//Only run when commanded to be in remote
q_stPump.xIlkOK := q_stPump.q_xRemoteDO AND q_stPump.i_xAlarmOK;

IF q_stPump.xIlkOK THEN
    q_stPump.q_xRunDO := q_stPump.pv_xRunSW;
    ELSE
        q_stPump.PV_xRunSW := FALSE;
        q_stPump.q_xRunDO := FALSE;
END_IF

q_stPump.xLspd_IlkENA := q_stPump.xIlkOK;

IF q_stPump.xLspd_IlkENA THEN
    q_stPump.q_xLspdDo := q_stPump.xLspdSW;
    ELSE
        q_stPump.xLspdSW := FALSE;
        q_stPump.q_xLspdDo := FALSE;
END_IF

//resetTmr (In := iq_stPump.xResetSW, PT := T#2S);
//IF resetTmr.Q THEN
//	iq_stPump.xResetSW := FALSE;
//END_IF

q_stPump.q_xResetDo := NOT q_stPump.i_xIsRun AND q_stPump.xResetSW;

//countdown Timer
TONtmr (IN := q_stPump.i_xIsRun, PT := T#20S);
q_stPump.RdyTmr := TO_REAL(TONtmr.PT) - TO_REAL(TONtmr.ET);

(*State evaluation*)
IF NOT q_stPump.i_xAlarmOK THEN
    q_stPump.eState := pumpFAULT;
ELSIF NOT q_stPump.q_xRunDo AND q_stPump.i_xAlarmOK THEN
        q_stPump.eState := pumpSTOPPED;
ELSIF q_stPump.q_xRunDo AND NOT q_stPump.i_xIsRun THEN
        q_stPump.eState := pumpSTARTING;
ELSIF q_stPump.i_xIsRun THEN
        q_stPump.eState := pumpRUNNING;
ELSE
    q_stPump.eState := pumpFAULT;
END_IF

//Mapping
M_IO();

METHOD M_Alarm : BOOL
VAR_INPUT
END_VAR
M_alarm := THIS^.q_stPump.i_xAlarmOK;   // 0 = no alarm | 1 = alarm
END_METHOD

METHOD M_AlarmOK : BOOL
VAR_INPUT
END_VAR
M_AlarmOK := THIS^.q_stPump.i_xAlarmOK;
END_METHOD

METHOD M_IO : BOOL
VAR_INPUT
END_VAR
(* Output *)
    q_xRunDO 	:= THIS^.q_stPump.q_xRunDO;
    q_xResetDo := THIS^.q_stPump.q_xResetDo;
    q_xLspdDo := THIS^.q_stPump.q_xLspdDo;
    q_xRemote := THIS^.q_stPump.q_xRemoteDo;
(* Input *)
    THIS^.q_stPump.i_xAlarmOK :=	THIS^.i_xAlarm;
    THIS^.q_stPump.i_xIsRun :=	THIS^.i_xIsRun;
END_METHOD

METHOD M_IsRun : BOOL
VAR_INPUT
END_VAR
M_IsRun := THIS^.q_stPump.i_xIsRun;
END_METHOD

METHOD M_Lspd : BOOL
VAR_INPUT
    lowspeed : BOOL;  // Set low speed setting
END_VAR
THIS^.q_stPump.xLspdSW := lowspeed;
END_METHOD

METHOD M_Remote : BOOL
VAR_INPUT
    remote : BOOL; // Remote command
END_VAR
this^.q_stPump.xRemoteSW := remote;
END_METHOD

METHOD M_Reset : BOOL
VAR_INPUT
    reset : BOOL; // Set true to clear faults
END_VAR
this^.q_stPump.xResetSW := reset;
END_METHOD

METHOD PUBLIC M_Run : BOOL
VAR_INPUT
    run:bool; // set to true to run, false to stop;
END_VAR

this^.q_stPump.pv_xRunSW := run;
END_METHOD

END_FUNCTION_BLOCK

// ---- POUs/Functions/Pumps/FB_PIP_Gamma_V2.TcPOU
(* This function block does basic controls FOR the ION pump connected to a Gamma QPCe controller. *)
{attribute 'reflection'}
FUNCTION_BLOCK FB_PIP_Gamma_V2 Extends FB_Pump
VAR_INPUT
END_VAR
VAR_OUTPUT
    {attribute 'pytmc' := '
    pv:
    '}
    stPump	:	ST_PIP; //Gamma Ion pump structure
    q_IG	:	ST_VG; //When ion pump is used as a measuring device for interlocking gate valves
END_VAR
VAR
    rPRESS : REAL;

    rV : REAL;

    (* IO Controls *)
    i_iPRESS  AT %I*: INT;  //
    i_xSP_DI  AT %I* : BOOL; // NO contact //function of relay set on the QPC to HV output state

    // For logging
    tPumpErrorTimeout : TON := (PT:=T#10S); // Timeout pump start if pressure < 1E-11 for more than 10s.

    {attribute 'instance-path'}
    {attribute 'noinit'}
    sPath: STRING;
    fbGetCurTaskIdx  : GETCURTASKINDEX;
    fbWritePersistentData           : WritePersistentData;

END_VAR
VAR CONSTANT
    rMaxPressure : REAL :=1E-4; // Default protection setpoint as per the gamma QPCe manual
    rMinPressure : REAL :=1E-11;
END_VAR
VAR PERSISTENT
END_VAR

(*Pump STATE*)
tPumpErrorTimeout(IN:=(q_IG.rPRESS <= rMinPressure AND stPump.i_xHV_DI));

IF q_IG.rPRESS <= rMinPressure AND stPump.i_xHV_DI THEN
    IF tPumpErrorTimeout.Q THEN
        stPump.eState := pumpFAULT;
        tPumpErrorTimeout(IN:=FALSE);
    END_IF
ELSIF q_IG.rPRESS <= rMinPressure AND NOT stPump.i_xHV_DI THEN
    stPump.eState := pumpSTOPPED;
ELSIF stPump.i_xHV_DI THEN
    stPump.eState := pumpRUNNING;
ELSE
    stPump.eState := pumpFAULT;
END_IF

(*Update output gauge values*)
ACT_SetGauge();
(*Soft IO Mapping*)
IO();
// Log States and triggers
ACT_Logger();

ACTION ACT_Logger:
//STATE Logger
IF ePrevState <> stPump.eState THEN
      CASE stPump.eState OF
        pumpFAULT:
            fbLogger(sMsg:='Pump Fault.', eSevr:=TcEventSeverity.Critical);
        pumpSTOPPED:
            fbLogger(sMsg:='Pump stopped.', eSevr:=TcEventSeverity.Critical);
        pumpRUNNING:
            fbLogger(sMsg:='Pump running.', eSevr:=TcEventSeverity.Info);
      END_CASE
      ePrevState := stPump.eState;
  END_IF
END_ACTION

ACTION ACT_SetGauge:
(*MG*)
(* convert the analog input into readable pressure*)
(* use logarithmic Pressure calculation, Output= Normal and Offset = 0*)
rV := 10*INT_TO_REAL(i_iPress)/32767;
//Manual Page 9

if (stPump.bOutputInverted) THEN
    rPRESS := LREAL_TO_REAL(EXPT(10,(rV-stPump.iOffset)*-1));
ELSE
    rPRESS := LREAL_TO_REAL(EXPT(10,(rV-stPump.iOffset)));
END_IF

q_IG.rPRESS := rPRESS;
stPump.rPRESS := rPRESS;

IF stPump.eState := pumpRUNNING THEN
    q_IG.xPRESS_OK := TRUE;
ELSE
    q_IG.xPRESS_OK := FALSE;
END_IF

q_IG.sPath := This^.stPump.sPath;
END_ACTION

ACTION IO:
stPump.xError := (stPump.eState = pumpFAULT);

(*inputs*)
stPump.i_iPRESS:=	i_iPRESS;
stPump.i_xHV_DI:=	i_xSP_DI;

 This^.stPump.sPath:= sPath;
END_ACTION

END_FUNCTION_BLOCK

// ---- POUs/Functions/Pumps/FB_PIP_SIP.TcPOU
(* This function block does basic controls FOR the ION pump connected to a SAES SIP controller.
 Provides interlocking interface. Enable HV only when interlock gauge press is less than 1.0E-4 Torr *)
{attribute 'reflection'}
FUNCTION_BLOCK FB_PIP_SIP Extends FB_Pump
VAR_INPUT
    i_stGauge	:	ST_VG; //Ion or Pirani gauge for pump interlock
    i_xOverrideMode : BOOL; (*To be linked to global override bit. This Overrides Vacuum interlock logic*)
END_VAR
VAR_OUTPUT
    {attribute 'pytmc' := '
    pv:
    '}
    stPump	:	ST_PIP; //Gamma Ion pump structure
    q_IG	:	ST_VG; //When ion pump is used as a measuring device for interlocking gate valves
END_VAR
VAR
 rPRESS : REAL;
 iTermBits: UINT := 32767 ; // The terminal's maximum value in bits
 rV : REAL;
 timer:TON;

 (* IO Controls *)
 q_xHVEna_DO AT %Q*: BOOL;	// Enable High Voltage when TRUE
 i_iPRESS  AT %I*: INT;  //
 i_xIP_ON  AT %I* : BOOL;
 i_xError  AT %I* : BOOL;

// For logging
tTimeOutAction : F_TRIG;
tOverrideActivated : R_TRIG;

tPumpStartTimeout : TON := (PT:=T#10s); // Timeout pump start if pressure < 1E-11 for more than 10s.
MinPressure : REAL:= 1E-11; // Minimum readback pressure, pump must register pressure above this to be considered running

//Overrides
    tonOvrd	:	TON;
    tonDelOK : TON;
    rtOK	:	R_TRIG;
    tOvrd	:	TIME := T#10s;

    {attribute 'instance-path'}
    {attribute 'noinit'}
    sPath: STRING;
END_VAR
VAR CONSTANT
     rDefaultHVEna_SP : REAL :=1E-4; // Default protection setpoint as per the gamma QPCe manual
END_VAR
VAR PERSISTENT
    rHVEna_SP : REAL;
END_VAR

(* Does Gamma Ion pump HV interlock. Enable HV only when interlock gauge press is less than 1.0E-4 Torr *)

(*Ensures the set point is not higher than 1.0E-4*)
IF (stPump.rHVEna_SP > rDefaultHVEna_SP) THEN
    stPump.rHVEna_SP := rDefaultHVEna_SP;
END_IF

(* Interlock *)
//stPump.xHV_ExtIlk  := i_stGauge.xPRESS_OK AND (i_stGauge.rPRESS <= stPump.rHVEna_SP);//AND NOT tPumpStartTimeout.Q); //ADP

(* Enable HV *)
IF i_stGauge.rPRESS <= stPump.rHVEna_SP AND i_stGauge.xPRESS_OK THEN
    IF (stPump.xAutoOn) AND NOT (stPump.q_xHVEna_DO) THEN  stPump.q_xHVEna_DO := TRUE;
    ELSE stPump.q_xHVEna_DO := stPump.xHVEna_SW OR ((tonOvrd.Q AND i_xOverrideMode));
    END_IF
    stPump.xILKOk:= TRUE;
ELSIF stPump.q_xHVEna_DO (*AND timer.Q*) THEN
    IF q_IG.rPRESS > (stPump.rHVEna_SP + stPump.rHYS_PR) THEN // Ion pumps when running switches off based on their own pressure readings
        stPump.q_xHVEna_DO := FALSE;
        stPump.xHVEna_SW := FALSE;
        stPump.xILKOk := FALSE;
    ELSE
        stPump.q_xHVEna_DO := stPump.xHVEna_SW OR ((tonOvrd.Q AND i_xOverrideMode));
    END_IF
ELSIF (tonOvrd.Q AND i_xOverrideMode) THEN
    stPump.q_xHVEna_DO := TRUE;
ELSE
    stPump.q_xHVEna_DO  := FALSE;
    stPump.xHVEna_SW := FALSE;
    stPump.xILKOk := FALSE;
END_IF


//stPump.q_xHVEna_DO := stPump.xHVEna_SW AND stPump.xHV_ExtIlk;
//stPump.xHVEna_SW := stPump.q_xHVEna_DO;

timer(IN:= NOT stPump.q_xHVEna_DO, PT:= T#1s);

// TAW Experimental ion pump timeout
tPumpStartTimeout(IN:=(NOT stPump.i_xHV_DI AND stPump.q_xHVEna_DO));
tTimeOutAction(CLK:=tPumpStartTimeout.Q);
IF tTimeOutAction.Q THEN  fbLogger(sMsg:='Pump time out.', eSevr:=TcEventSeverity.Critical); END_IF



(*Pump STATE*)
IF tPumpStartTimeout.Q OR i_xError  THEN //Pump timeout
    stPump.eState := pumpFAULT;
ELSIF stPump.q_xHVEna_DO AND NOT stPump.i_xHV_DI THEN
    stPump.eState := pumpSTARTING;
ELSIF NOT stPump.q_xHVEna_DO AND NOT stPump.i_xHV_DI THEN
    stPump.eState := pumpSTOPPED;
ELSIF stPump.q_xHVEna_DO AND stPump.i_xHV_DI THEN
    stPump.eState := pumpRUNNING;
ELSIF NOT stPump.q_xHVEna_DO AND stPump.i_xHV_DI THEN
    stPump.eState := pumpSTOPPING;
ELSE
    stPump.eState := pumpFAULT;
END_IF



(*Update output gauge values*)
ACT_SetGauge();
(*Soft IO Mapping*)
IO();
ACT_IlkOverride();
// Log States and triggers
ACT_Logger();
(*Load or save the persistent variables*)
ACT_Persistent();

ACTION ACT_IlkOverride:
(* Override logic *)
(* Goal: give ability to override, but do so in a way that people won't forget it.
Solution: Override only after ten seconds of override, protect against blips,
when the Pump permission goes true for more than ten seconds consistently, remove override
*)

tonDelOK(IN:=stPump.xILKOk, PT:=T#10S);
rtOK(CLK:=tonDelOK.Q);
IF rtOK.Q AND stPump.pv_xOvrdStart THEN
    stPump.pv_xOvrdStart :=FALSE;
    if (stPump.eState = pumpRUNNING) AND (i_xOverrideMode) THEN stPump.xHVEna_SW:= TRUE; END_IF
    //Log
    fbLogger(sMsg:='Override expired', eSevr:=TcEventSeverity.Warning);
END_IF
// Release the Force DO bit when the system override is false
IF NOT(i_xOverrideMode) THEN stPump.pv_xOvrdStart :=FALSE; END_IF
//Override timer
tonOvrd(IN:= stPump.pv_xOvrdStart, PT:=tOvrd);
END_ACTION

ACTION ACT_Logger:
// ILK logger

IF NOT (stPump.xILKOk) AND ((ePrevState = pumpRUNNING) OR (ePrevState = pumpSTARTING)) AND NOT tonOvrd.Q THEN
    fbLogger(sMsg:='Pump turned off due to loss of interlock.', eSevr:=TcEventSeverity.Critical);
END_IF

//STATE Logger
IF ePrevState <> stPump.eState THEN
      CASE stPump.eState OF
        pumpFAULT:
            fbLogger(sMsg:='Pump Fault.', eSevr:=TcEventSeverity.Critical);
          pumpSTOPPED:
            fbLogger(sMsg:='Pump stopped.', eSevr:=TcEventSeverity.Critical);
        pumpSTARTING:
            fbLogger(sMsg:='Pump starting.', eSevr:=TcEventSeverity.Info);
        pumpRUNNING:
            fbLogger(sMsg:='Pump running.', eSevr:=TcEventSeverity.Info);
        pumpSTOPPING:
            fbLogger(sMsg:='Pump stopping.', eSevr:=TcEventSeverity.Info);
      END_CASE
      ePrevState := stPump.eState;
  END_IF


  // Log Action
tAction(CLK:=  stPump.q_xHVEna_DO);
IF tAction.Q THEN fbLogger(sMsg:='Pump commanded to start', eSevr:=TcEventSeverity.Info); END_IF
// Log override mode enabled
tOverrideActivated(CLK:= (tonOvrd.Q AND i_xOverrideMode));
IF tOverrideActivated.Q THEN fbLogger(sMsg:='Pump override mode activated', eSevr:=TcEventSeverity.Warning); END_IF


// Log FAULT
tFault(CLK:=  NOT tPumpStartTimeout.Q);
IF tFault.Q THEN fbLogger(sMsg:='Pump Fault', eSevr:=TcEventSeverity.Critical); END_IF
END_ACTION

ACTION ACT_Persistent:
(*On first PLC pass, load the persistent value into the structrue variable*)
IF (SUPER^.bRestorePersistentData) THEN
    SUPER^.bRestorePersistentData	:= FALSE;
    IF (rHVEna_SP <> 0) THEN
        stPump.rHVEna_SP := rHVEna_SP;
    END_IF;
END_IF
(*Check if a new value has been written in the structure variable copy it to the persistent variable*)
IF NOT (stPump.rHVEna_SP = rHVEna_SP) THEN
    rHVEna_SP := stPump.rHVEna_SP;
END_IF;
END_ACTION

ACTION ACT_SetGauge:
(*MG*)
(* convert the analog input into readable pressure*)
(* use logarithmic Pressure calculation, Output= Normal and Offset = 0*)
If (iTermBits=0) THEN iTermBits := 32767;END_IF
rV := 10*INT_TO_REAL(i_iPress)/iTermBits;
//Manual Page 29
IF (rV >= 2.5) THEN
    rPRESS := LREAL_TO_REAL((0.000000001*EXP(1.8421*rV))/65);
    ELSE
    rPRESS := LREAL_TO_REAL((0.0000000008*EXP(1.9315*rV))/65);
END_IF
// Min. measured pressure
IF (rPRESS < 1E-11) AND NOT (rPRESS = 0)  THEN
    rPRESS := 1E-11;
END_IF

IF (stPump.q_xHVEna_DO) THEN
    q_IG.rPRESS := rPRESS;
    stPump.rPRESS := rPRESS;
END_IF


IF (stPump.i_xHV_DI) AND (q_IG.rPRESS < q_IG.rVAC_SP) THEN //ADP// AND (q_IG.rPRESS<>0) AND stPump.q_xHVEna_DO) THEN
    q_IG.xPRESS_OK := TRUE;
    ELSE
    q_IG.xPRESS_OK := FALSE;
END_IF

q_IG.sPath := This^.stPump.sPath;
END_ACTION

ACTION IO:
stPump.sIlkDeviceName := This^.i_stGauge.sPath;
stPump.xError := i_xError;// (stPump.eState = pumpFAULT);
stPump.xOverrideMode := i_xOverrideMode;
(*inputs*)
stPump.i_iPRESS:=	i_iPRESS;
stPump.i_xHV_DI:=	i_xIP_ON;
(*output*)
q_xHVEna_DO:=  stPump.q_xHVEna_DO; //According to Manual pin should be grounded to activate function

 This^.stPump.sPath:= sPath;
END_ACTION

METHOD M_AutoOn : BOOL
VAR_INPUT
END_VAR
this^.stPump.xAutoOn:= TRUE; // Pump is set to auto start when the pressure is low enough
END_METHOD


METHOD PUBLIC M_Run : BOOL
VAR_INPUT
    run:bool; // set to true to run, false to stop;
END_VAR

this^.stPump.xHVEna_SW := run;
END_METHOD

END_FUNCTION_BLOCK

// ---- POUs/Functions/Pumps/FB_PTM_Agilent.TcPOU
(* This function block does basic controls FOR the Agilent TV Turbo pump. Turns off pump
in the event of errors/ warnings. Provides interlocking interface.*)
FUNCTION_BLOCK FB_PTM_Agilent EXTENDS FB_Pump
VAR_IN_OUT

END_VAR
VAR_INPUT
    i_xExtILKOk : BOOL; // Connect to external interlock logic(e.g TURBO_ILK Function), TRUE if not used.
    i_stGauge	:	ST_VG; //Pirani backing gauge for pump interlock
    i_rMaxBackingPressure : REAL;
END_VAR
VAR_OUTPUT
    {attribute 'pytmc' :=' pv:'}
    iq_stPtm	:	ST_AgilentPTM;

END_VAR
VAR
    {attribute 'instance-path'}
    {attribute 'noinit'}
    sPath: STRING;
    //xRunOk	:	BOOL;
    nMaxR1Fault: INT :=5;
    nR1Fault : INT;
    tFaultWindowDuration : TIME := T#300S;
    tR1FaultDuration : TIME := T#120S;
    tTimeOutDuration: TIME:= T#10M;
    tFaultWindowElapsed: TON;
    tR1Fault : TON;
    tStartTimeOut : TON;
    tR1TimeOut: TON;
    step : INT :=0;
    nErrorCode: INT :=0;
    xBackingPressureOK: BOOL;
    iMaxSpeed : INT:=963;

    rPowerScale: REAL:=10;//W
    rCurrentScale: REAL:=1;//A

    (*I/Os*)
    i_xSTART 	AT%I*:	BOOL;
    i_xR1	AT%I*	:  BOOL;
    i_xR2	AT%I*	:  BOOL;
    i_xLSpd	AT%I*:  BOOL;
    i_iTempMon AT%I*: INT;
    i_iPowerMon AT%I*: INT;
    i_iCurrentMon AT%I*: INT;
    i_iRawSpeed AT %I* : INT;
    i_xFault AT%I*	:	BOOL;
    q_RunDO AT%Q*	:	BOOL;
    q_xLSpd	AT%Q*	:  BOOL;


    // For logging
  //  Msg : FB_FormatString;
   // fbJson : FB_JsonSaxWriter;
   tOverrideActivated : R_TRIG;

    iTermBits: UINT := 32767 ; // The terminal's maximum value in bits
END_VAR

(* Basic Agilent Turbo Controls *)
(* M. Ghaly, 2018-9-26 *)

(*connect External interlock to structure variable*)
//iq_stPtm.xExtRunOk := i_xExtILKOk;

(* state machine *)
CASE (step) OF
(*Pump Stopped State*)
    0: // Pump Stopped State
        iq_stPtm.xRunSW:=FALSE;
        //Reset Output signals;
        iq_stPtm.q_RunDO:=FALSE;
        iq_stPtm.q_xSS := FALSE;
        iq_stPtm.q_xLSpd:= FALSE;
        //Reset timer
        tFaultWindowElapsed.IN := FALSE;
        nR1Fault := 0;
        iq_stPtm.eState := pumpSTOPPED;
        step :=10;

(*Idle State waiting to start*)
    10: // Idle State, waiting for the xRunSwitch
        IF iq_stPtm.xExtRunOk  AND iq_stPTM.xRunSW THEN
            iq_stPtm.q_RunDO := iq_stPTM.xRunSW; //
            step:=20;
        END_IF
(*Pump Starting State*)
    20: // Pump is starting
        nErrorCode:=0;
        iq_stPtm.q_RunDO := iq_stPTM.xRunSW; // done in previous state
        IF (*(NOT iq_stPtm.i_xR1) AND*)iq_stPtm.i_xSTART  THEN
        iq_stPtm.eState := pumpSTARTING;
        step:= 40;
        ELSIF tStartTimeOut.Q THEN
            step:=90; // or fault state
            nErrorCode:=950;
        END_IF
        // should check R1 ?? check Fault condition?


    40: // Pump is starting
        iq_stPtm.eState := pumpSTARTING;
        IF   NOT iq_stPtm.i_xR1 AND NOT iq_stPtm.i_xSTART  THEN
            step := 0 ;
        ELSIF NOT iq_stPtm.i_xR1 AND iq_stPtm.i_xSTART  THEN
            step :=40;
        ELSIF iq_stPtm.i_xR1 AND NOT iq_stPtm.i_xSTART THEN
            step:= 50;
        END_IF
        IF tR1TimeOut.Q THEN
            step:= 90;
            iq_stPtm.xPumpFaultLock := TRUE;
            nErrorCode:= 930; // R1 Signal at Start time out.
           // fbLogger(sMsg:='Timeout: Pump could not achieve running speed.', eSevr:=TcEventSeverity.Warning);
        END_IF

    50: // Pump is Running (Normal Operation) ( R1 is True and STARTing is FALSE)
        iq_stPtm.eState := pumpRUNNING;
        IF NOT iq_stPtm.i_xR1 THEN
            nR1Fault:= nR1Fault+1 ;
            tFaultWindowElapsed.IN := TRUE; ///
            //tR1Fault.IN := TRUE;
            step :=60;
        END_IF

        //Log new state
        IF ePrevState <> iq_stPtm.eState THEN
            //fbLogger(sMsg:='Pump at speed.', eSevr:=TcEventSeverity.Verbose);
            ePrevState := iq_stPtm.eState;
        END_IF

    60: // Pump is Running (Not Nomral Operation) (R1 is False, pump not @ speed )
        IF ((nR1Fault = nMaxR1Fault) AND NOT tFaultWindowElapsed.Q) OR (tR1Fault.Q) THEN // number of fault occured during the same time window
            step:= 90;
            tR1Fault.IN := FALSE;
            tFaultWindowElapsed.IN := FALSE;
            iq_stPtm.xPumpFaultLock := TRUE;
            nErrorCode:= 920; // R1 Signal Lost multiple times.
            //fbLogger(sMsg:='Running signal Lost multiple times.', eSevr:=TcEventSeverity.Warning);
        ELSIF tFaultWindowElapsed.Q  THEN
            tFaultWindowElapsed.IN := FALSE;
            nR1Fault := 0;
        ELSIF iq_stPtm.i_xR1 THEN
            tR1Fault.IN := FALSE;
            step:=50;
        END_IF

    90: // Pump Fault STATE
        iq_stPtm.xRunSW:=FALSE;
        iq_stPtm.q_RunDO:=FALSE;
        iq_stPtm.q_xSS := FALSE;
        iq_stPtm.q_xLSpd:= FALSE;
        iq_stPtm.eState := pumpFAULT;
        step := 95;

    95:
        IF (NOT iq_stPtm.xPumpFaultLock) OR iq_stPtm.xRunSW THEN
            step:=0;
        END_IF
END_CASE

(* Interrupts *)
(* FAULT signal*)
IF (iq_stPtm.i_xFault) AND (step < 90 ) THEN
    iq_stPtm.eState := pumpFAULT; // no need taken care of in the state
    iq_stPtm.xPumpFaultLock := TRUE;
    nErrorCode := 900; // Pump Controller FAULT
    step:=90;
END_IF


(*Pump Lock Reset bit*)
IF (iq_stPtm.xResetSW ) THEN
    iq_stPtm.xResetSW := FALSE;
    iq_stPtm.xPumpFaultLock := FALSE;
END_IF

(*Check backing gauge pressure*)
//xBackingPressureOK := i_stGauge.xPRESS_OK AND ( i_stGauge.rPRESS < iq_stPtm.rBackingPressureSP);

(* Interlock Sum *)
iq_stPtm.xExtRunOk := i_xExtILKOk AND NOT iq_stPtm.i_xFault AND NOT iq_stPtm.xPumpFaultLock AND NOT(tILK.Q);

IF NOT iq_stPtm.xExtRunOk AND (NOT (step >= 90)) THEN
    step:=0;
END_IF

(*Stop By the Operator and not due to fault *)
IF (NOT iq_stPtm.xRunSW) AND (NOT (step >= 90)) AND (NOT (step = 10)) THEN
    step := 0;
END_IF

// Log faults Moved to ACT_Logger
(*tErrorPresent(CLK:=iq_stPtm.xPumpFaultLock);
IF tErrorPresent.Q THEN
    fbJson.StartObject();
    fbJson.AddKey('vacuum_typecode');
    fbJson.AddUdint(nErrorCode);
    fbJson.EndObject();
    fbLogger.sJson := fbJson.GetDocument();
    fbLogger(sMsg:='Turbo control fault', eSevr:=TcEventSeverity.Warning);
    fbJson.ResetDocument();
END_IF
*)

(* Timers *)
tFaultWindowElapsed(PT:=tFaultWindowDuration);
tR1Fault(IN:= (step = 60), PT:=tR1FaultDuration);
tStartTimeOut(IN := (step=20), PT:=tTimeOutDuration);
tR1TimeOut(IN := (step=40), PT:=tTimeOutDuration);
(* IO Mapping*)
IO();
(*Assign Error Message*)
iq_stPtm.sError := ErrorMessage(nErrorCode, iq_stPtm.eState);
// Log States and triggers
ACT_Logger();
(*Validate Backing Pressure set point doesn't exceed the Maximum backingPressure*)
iq_stPtm.rBackingPressureSP := BackingPressureSetPoint(iq_stPtm.rBackingPressureSP,i_rMaxBackingPressure);
ACT_Interlock();
(*Load or save the persistent variables*)
ACT_Persistent();

ACTION ACT_Interlock:
This^.tILK(IN:= (i_stGauge.rPRESS>=iq_stPtm.rBackingPressureSP), PT:=T#5S, Q=> );
END_ACTION

ACTION ACT_Logger:
//STATE Logger
// ILK logger
IF NOT i_xExtIlkOK AND ePrevState = pumpRUNNING THEN
         fbLogger(sMsg:='Lost external interlock while pump was running.', eSevr:=TcEventSeverity.Critical);
END_IF


IF ePrevState <> iq_stPTM.eState THEN
      CASE iq_stPTM.eState OF
        pumpFAULT:
            fbLogger(sMsg:='Pump Fault.', eSevr:=TcEventSeverity.Critical);
          pumpSTOPPED:
            fbLogger(sMsg:='Pump stopped.', eSevr:=TcEventSeverity.Critical);
        pumpSTARTING:
            fbLogger(sMsg:='Pump starting.', eSevr:=TcEventSeverity.Info);
        pumpRUNNING:
            fbLogger(sMsg:='Pump running.', eSevr:=TcEventSeverity.Info);
      END_CASE
      ePrevState := iq_stPTM.eState;
  END_IF

// Log Action
tAction(CLK:=  iq_stPTM.q_RunDO);
IF tAction.Q THEN fbLogger(sMsg:='Pump commanded to start', eSevr:=TcEventSeverity.Info); END_IF


// Log FAULT
tFault(CLK:= iq_stPTM.i_xFault OR iq_stPtm.xPumpFaultLock);
IF tFault.Q THEN fbLogger(sMsg:=iq_stPtm.sError, eSevr:=TcEventSeverity.Critical); END_IF
END_ACTION

ACTION ACT_Persistent:
(*On first PLC pass, load the persistent value into the structrue variable*)
IF (SUPER^.bRestorePersistentData) THEN
    SUPER^.bRestorePersistentData	:= FALSE;
    IF (rBackingPressureSP <> 0) THEN
        iq_stPTM.rBackingPressureSP := rBackingPressureSP;
    END_IF;
    IF (rInletPressureSP <> 0) THEN
        iq_stPTM.rInletPressureSP := rInletPressureSP;
    END_IF;
END_IF
(*Check if a new value has been written in the structure variable copy it to the persistent variable*)
IF NOT (iq_stPTM.rBackingPressureSP = rBackingPressureSP) THEN
    rBackingPressureSP:= iq_stPTM.rBackingPressureSP;
END_IF;

IF NOT (iq_stPTM.rInletPressureSP = rInletPressureSP) THEN
    rInletPressureSP := iq_stPTM.rInletPressureSP;
END_IF;
END_ACTION

METHOD BackingPressureSetPoint : REAL
VAR_INPUT
    i_SetPoint : REAL;
    rMaxBackingPressure: REAL;
END_VAR
BackingPressureSetPoint := Min(i_SetPoint , rMaxBackingPressure);
END_METHOD

METHOD PUBLIC ErrorMessage : STRING
VAR_INPUT
    nErrorCode : INT;
    eState: E_PumpState;
END_VAR
IF (eState = pumpFAULT ) THEN
    CASE nErrorCode OF
        950:
            ErrorMessage := 'Pump Starting Fault';
        930:
            ErrorMessage := 'Pump could not achieve running speed';

        920:
            ErrorMessage := 'Running at speed signal lost multiple times';

        900:
            ErrorMessage := 'Pump Controller Fault';
    END_CASE

END_IF
END_METHOD

ACTION IO:
(*inputs*)
iq_stPtm.i_xSTART:=	i_xSTART;
iq_stPtm.i_xR1:=	i_xR1;
iq_stPtm.i_xR2:=	i_xR2;
iq_stPtm.i_xLSpd:=	i_xLSpd;
iq_stPtm.i_xFault:=	i_xFault;
(* Real-value calculation *)
If (iTermBits=0) THEN iTermBits := 32767;END_IF
iq_stPtm.i_rCurrentMon := (10*INT_TO_REAL(i_iCurrentMon)/iTermBits)*rCurrentScale;
iq_stPtm.i_rTempMon := 10*INT_TO_REAL(i_iTempMon)/iTermBits;
iq_stPtm.i_rPowerMon := (10*INT_TO_REAL(i_iPowerMon)/iTermBits)*rPowerScale;
iq_stPtm.i_diCurSpd := 10*LREAL_TO_DINT(INT_TO_REAL(i_iRawSpeed)/iTermBits);


(*outputs*)
q_RunDO := iq_stPtm.q_RunDO;
q_xLSpd := iq_stPtm.q_xLSpd;
END_ACTION

METHOD PUBLIC M_Run : BOOL
VAR_INPUT
    run:bool; // set to true to run, false to stop;
END_VAR

this^.iq_stPtm.xRunSW := run;
END_METHOD

METHOD M_SetBits : BOOL
VAR_INPUT
    TermBits : UINT; // The terminal's maximum value in bits
END_VAR
This^.iTermBits := TermBits;
END_METHOD

METHOD M_SetCurrentScale : BOOL
VAR_INPUT
    Scale:REAL;//In Amps
END_VAR
This^.rCurrentScale := Scale;
END_METHOD

METHOD M_SetMaxSpeed : BOOL
VAR_INPUT
    iMaxSpeed: INT; //963Hz for 3.1,300HT and 1010Hz for 401 and 1350 for 81
END_VAR
this^.iMaxSpeed := iMaxSpeed;
END_METHOD

METHOD M_SetPowerScale : BOOL
VAR_INPUT
    Scale:REAL;//In Watt
END_VAR
This^.rPowerScale := Scale;
END_METHOD

METHOD PUBLIC M_TurboIsOn : BOOL
VAR_INPUT
END_VAR
M_TurboIsOn := (This^.iq_stPtm.eState =  E_PumpState.pumpSTARTING ) OR (This^.iq_stPtm.eState =  E_PumpState.pumpRUNNING );
END_METHOD

END_FUNCTION_BLOCK

// ---- POUs/Functions/Pumps/FB_PTM_Ebara_011M.TcPOU
(* This function block does basic controls FOR the Ebara Turbo pump connected to the ETC011M Controller.
 Turns off pump in the event of errors/ warnings. Provides interlocking interface.*)
{attribute 'no_check'}
FUNCTION_BLOCK FB_PTM_Ebara_011M EXTENDS FB_Pump
VAR_IN_OUT
END_VAR
VAR_INPUT
    i_rMaxBackingPressure : REAL := 3;
    i_iMinSpeed : DINT := 100; //check pump manual for setting
    i_iMaxSpeed : DINT := 560; // check pump manual for setting
    i_xExtILKOk : BOOL; // Connect to external interlock logic, TRUE if not used.
END_VAR
VAR_OUTPUT
    {attribute 'pytmc' := '
    pv:
    '}
    iq_stPTM : ST_EbaraPTM;
END_VAR
VAR
    TOF_SetSpeed: TON := (PT:=T#1S);
    TOF_RESET: TON :=(PT:=T#1S);
    i_iADCBits : UINT := 12;
    (*IO*)
    (*inputs*)
    i_xDecel AT %I* : BOOL; //Link to brake input
    i_xAccel AT %I* : BOOL;
    i_xRotate AT %I* : BOOL;
    i_xFaultNC AT %I* : BOOL;// remove?
    i_xAtSpd AT %I* : BOOL;
    i_iRawSpeed AT %I* : INT; // Link to Analog input

    (*output*)
    q_xStart AT %Q* : BOOL; // link to output
    q_xStop AT %Q* : BOOL; //Link to output
    q_xReset AT %Q* : BOOL;
    q_xProtection AT %Q* : BOOL;
    q_xSetSpeed AT %Q* : BOOL;
    q_iSpeedSet AT %Q* :INT;	//Link to analog Output


END_VAR

(* Ebara ETC control FB
Scott Stubbs & Alex W.
Modified Nov 2018 by M. Ghaly
*)

(* Switch processing *)
//TOF_START.IN := iq_stPTM.i_xStart;
//TOF_START();
//TOF_STOP.IN  := iq_stPTM.i_xStop;
//TOF_STOP();
//TOF_RESET.IN := iq_stPTM.i_xReset;
//TOF_RESET();

(* Simple protection reset *)
iq_stPtm.xExtRunOk:= i_xExtILKOk;
iq_stPTM.q_xProtection := TRUE;//iq_stPTM.xExtRunOk;

(*soft IO mapping*)
ACT_IO();

(* Basic pump supervisory section *)
    (* If override mode, ignore everything else *)
IF iq_stPTM.i_xOverride THEN
    IF iq_stPTM.xRunSW THEN
        iq_stPTM.q_RunDO:=TRUE;
    ELSE
        iq_stPTM.q_RunDO:=FALSE;
    END_IF
    //Handle faults - the way the Ebara cable is done, xFault is normally closed
ELSIF iq_stPTM.i_xFault OR (iq_stPTM.q_RunDO AND NOT iq_stPTM.xExtRunOk) THEN
    iq_stPTM.q_RunDO:=FALSE;
    //iq_stPTM.q_xProtection:=FALSE;
    iq_stPTM.xRunSW:=FALSE;
    //And one for when we need to start the pump normally. Only allows pump to be started if ILK ok.
ELSIF iq_stPTM.xRunSW AND iq_stPTM.xExtRunOk THEN
    iq_stPTM.q_RunDO:=TRUE;
END_IF
//One section for when pump is told to stop
IF NOT iq_stPTM.xRunSW THEN
        iq_stPTM.q_RunDO:=FALSE;
        IF (NOT iq_stPTM.i_xFault) AND (NOT iq_stPTM.i_xALARM) THEN iq_stPTM.eState := pumpSTOPPED; END_IF;
END_IF

//Set the Start and Stop outputs to Run do . check manual.
iq_stPTM.q_xStart := iq_stPTM.q_xStop := iq_stPTM.q_RunDO;

(* to reset the Input speed OK bit *)
 TOF_SetSpeed (IN:= iq_stPTM.iq_xSpeedSet, Q => );
 IF TOF_SetSpeed.Q THEN iq_stPTM.iq_xSpeedSet:= FALSE;
 END_IF
 (* to reset the Reset Bit *)
 IF (iq_stPTM.xResetSW ) THEN  iq_stPTM.q_xReset := TRUE;
 END_IF
 TOF_RESET (IN:= iq_stPTM.q_xReset, Q => );
 IF TOF_RESET.Q THEN
    iq_stPTM.q_xReset:= FALSE;
    iq_stPTM.xResetSW := FALSE;
 END_IF


 (*Pump STATE*)
IF iq_stPtm.i_xFault THEN
    iq_stPtm.eState := pumpFAULT;
ELSIF iq_stPTM.i_xDecel AND NOT iq_stPtm.q_RunDO THEN
    iq_stPtm.eState := pumpSTOPPING;
ELSIF NOT iq_stPtm.q_RunDO AND NOT iq_stPTM.i_xFault THEN
    iq_stPtm.eState := pumpSTOPPED;
ELSIF NOT iq_stPtm.i_xAtSpd  AND iq_stPtm.q_RunDO THEN
    iq_stPtm.eState := pumpSTARTING;
ELSIF iq_stPtm.i_xAtSpd AND iq_stPtm.q_RunDO THEN
    iq_stPtm.eState := pumpRUNNING;
ELSE
    iq_stPtm.eState := pumpFAULT;
END_IF

(*Validate Backing Pressure set point doesn't exceed the Maximum backingPressure*)
iq_stPtm.rBackingPressureSP := BackingPressureSetPoint(iq_stPtm.rBackingPressureSP,i_rMaxBackingPressure);


(*soft IO mapping*)
ACT_IO();
// Log States and triggers
ACT_Logger();
(*Load or save the persistent variables*)
ACT_Persistent();

ACTION ACT_IO:
(*soft io mapping*)
(*inputs*)
    iq_stPTM.i_xDecel := i_xDecel ;
    iq_stPTM.i_xAccel :=	i_xAccel ;
    iq_stPTM.i_xRotate :=	i_xRotate;
    iq_stPTM.i_xNCFault :=	i_xFaultNC ;
    iq_stPTM.i_xAtSpd := i_xAtSpd;
    //iq_stPTM.i_iRawSpeed :=	i_iRawSpeed;
//V (AI/32767*10) * (33600 {Max RPM} - 100) / 5
(*outputs*)
    q_xStart:= iq_stPTM.q_xStart;
    q_xStop := iq_stPTM.q_xStop;
    q_xReset := iq_stPTM.q_xReset;
    q_xProtection := iq_stPTM.q_xProtection;
    q_xSetSpeed := iq_stPTM.iq_xSpeedSet;
(*Validate Set Speed within range *)
IF iq_stPTM.q_iSpeedSet  >= i_iMinSpeed AND iq_stPTM.q_iSpeedSet  <=i_iMaxSpeed THEN
    q_iSpeedSet  := LIMIT(0, DINT_TO_INT((iq_stPTM.q_iSpeedSet - i_iMinSpeed) / i_iMaxSpeed *16383/5),16383); //Max output 5V
    //:= DINT_TO_INT((iq_stPTM.q_iSpeedSet-100) / 33600 *32767/2); //Max 5V
END_IF

(* Pump speed calculation *)
iq_stPTM.i_diCurSpd := LREAL_TO_DINT(560*LREAL_TO_DINT(i_iRawSpeed)/16383);//(560*(INT_TO_REAL(i_iRawSpeed)/16383));// Manual page 28 (DC 0 to 5V -> 100 to 560Hz Rated Rotational Speed )
(*IF i_iRawSpeed / (EXPT(2,i_iADCBits)-1) * 10 >= 0.2 THEN //Speed reading appears zero at ~0.16V
iq_stPTM.i_diCurSpd := LREAL_TO_DINT(560*LREAL_TO_DINT(i_iRawSpeed)/16383);
//iq_stPTM.i_diCurSpd := LREAL_TO_DINT(i_iRawSpeed/(EXPT(2,i_iADCBits)-1)*67000);
//V (AI/(2^{# ADC bits} -1 ) * 10[ADC 10V scaling]) * (33600 [Max RPM] - 100) / 5
ELSE
    iq_stPTM.i_diCurSpd := 0;
END_IF*)

//Normally closed fault handling
iq_stPTM.i_xFault := NOT iq_stPTM.i_xNCFault; //??
END_ACTION

ACTION ACT_Logger:
//STATE Logger
IF NOT i_xExtIlkOK AND ePrevState = pumpRUNNING THEN
         fbLogger(sMsg:='Lost external interlock while pump was running.', eSevr:=TcEventSeverity.Critical);
END_IF


IF ePrevState <> iq_stPTM.eState THEN
      CASE iq_stPTM.eState OF
        pumpFAULT:
            fbLogger(sMsg:='Pump Fault.', eSevr:=TcEventSeverity.Critical);
          pumpSTOPPED:
            fbLogger(sMsg:='Pump stopped.', eSevr:=TcEventSeverity.Critical);
        pumpSTARTING:
            fbLogger(sMsg:='Pump starting.', eSevr:=TcEventSeverity.Info);
        pumpRUNNING:
            fbLogger(sMsg:='Pump running.', eSevr:=TcEventSeverity.Info);
        pumpSTOPPING:
            fbLogger(sMsg:='Pump decelerating.', eSevr:=TcEventSeverity.Info);
      END_CASE
      ePrevState := iq_stPTM.eState;
  END_IF

// ILK logger



// Log Action
tAction(CLK:=  iq_stPTM.q_RunDO);
IF tAction.Q THEN fbLogger(sMsg:='Pump commanded to start', eSevr:=TcEventSeverity.Info); END_IF


// Log FAULT
tFault(CLK:= iq_stPTM.i_xNCFault);
IF tFault.Q THEN fbLogger(sMsg:='Pump Lost Alarm OK bit', eSevr:=TcEventSeverity.Critical); END_IF
END_ACTION

ACTION ACT_Persistent:
(*On first PLC pass, load the persistent value into the structrue variable*)
IF (SUPER^.bRestorePersistentData) THEN
    SUPER^.bRestorePersistentData	:= FALSE;
    IF (rBackingPressureSP <> 0) THEN
        iq_stPTM.rBackingPressureSP := rBackingPressureSP;
    END_IF;
    IF (rInletPressureSP <> 0) THEN
        iq_stPTM.rInletPressureSP := rInletPressureSP;
    END_IF;
END_IF
(*Check if a new value has been written in the structure variable copy it to the persistent variable*)
IF NOT (iq_stPTM.rBackingPressureSP = rBackingPressureSP) THEN
    rBackingPressureSP:= iq_stPTM.rBackingPressureSP;
END_IF;

IF NOT (iq_stPTM.rInletPressureSP = rInletPressureSP) THEN
    rInletPressureSP := iq_stPTM.rInletPressureSP;
END_IF;
END_ACTION

METHOD PUBLIC BackingPressureSetPoint : REAL
VAR_INPUT
    i_SetPoint : REAL;
    rMaxBackingPressure: REAL;
END_VAR
BackingPressureSetPoint := Min(i_SetPoint , rMaxBackingPressure);
END_METHOD

METHOD PUBLIC M_Run : BOOL
VAR_INPUT
    run:bool; // set to true to run, false to stop;
END_VAR

this^.iq_stPtm.xRunSW := run;
END_METHOD

END_FUNCTION_BLOCK

// ---- POUs/Functions/Pumps/FB_PTM_MagDriveDigital.TcPOU
(* This function block does basic controls FOR the Leybold connected to the MagDriveDigital Controller.
 Turns off pump in the event of errors/ warnings. Provides interlocking interface.*)
FUNCTION_BLOCK FB_PTM_MagDriveDigital EXTENDS FB_Pump
VAR_IN_OUT

END_VAR
VAR_INPUT

    i_xExtILKOk : BOOL; // Connect to external interlock logic, TRUE if not used.
END_VAR
VAR_OUTPUT
{attribute 'pytmc' := '
    pv:
    '}
    iq_stPtm	:	ST_LeyboldPTM;
END_VAR
VAR
    xRunOk	:	BOOL;
    tofRemoteDelay	:	TOF;


    (*IO*)
    i_xAtSpd AT%I*: BOOL; // Normaml operation when true
    i_xFault AT%I*: BOOL; // Error NC
    i_xAccel AT%I*: BOOL;
     i_xDecel AT%I*: BOOL;
     i_xWarn AT%I*: BOOL;

    q_RunDO AT%Q*: BOOL; // Start/Stop
    q_xRemote AT%Q*: BOOL;
END_VAR

(* Basic MagDrive Digital Turbo Controls *)
(* A. Wallace, 2015-7-15 *)

tofRemoteDelay(IN:=iq_stPtm.q_RunDO, PT:=T#5S);

iq_stPtm.q_xRemote := tofRemoteDelay.Q;

(* Interlock Sum *)
iq_stPtm.xExtRunOk:= i_xExtILKOk;
xRunOk := iq_stPtm.xExtRunOk AND NOT iq_stPtm.i_xFault;

(* Basic pump supervisory section *)
IF xRunOk THEN
    iq_stPtm.q_RunDO := iq_stPTM.xRunSW;
ELSE
    iq_stPtm.xRunSW:=FALSE;
    iq_stPtm.q_RunDO:=FALSE;
END_IF

(*Pump STATE*)
IF iq_stPtm.i_xFault THEN
    iq_stPtm.eState := pumpFAULT;
ELSIF iq_stPTM.i_xDecel AND NOT iq_stPtm.q_RunDO THEN
    iq_stPtm.eState := pumpSTOPPING;
ELSIF NOT iq_stPtm.q_RunDO AND NOT iq_stPTM.i_xFault THEN
    iq_stPtm.eState := pumpSTOPPED;
ELSIF NOT iq_stPtm.i_xAtSpd  AND iq_stPtm.q_RunDO AND iq_stPTM.i_xAccel THEN
    iq_stPtm.eState := pumpSTARTING;
ELSIF iq_stPtm.i_xAtSpd AND iq_stPtm.q_RunDO THEN
    iq_stPtm.eState := pumpRUNNING;
ELSE
    iq_stPtm.eState := pumpFAULT;
END_IF


(*I/O soft mapping*)
ACT_IO();
// Log States and triggers
ACT_Logger();
(*Load or save the persistent variables*)
ACT_Persistent();

ACTION ACT_IO:
(*Inputs*)
iq_stPtm.i_xAtSpd := i_xAtSpd;
iq_stPtm.i_xFault := NOT i_xFault;
iq_stPtm.i_xAccel := i_xAccel;
iq_stPtm.i_xDecel := i_xDecel;
iq_stPtm.i_xWarn := i_xWarn;

(*Outputs*)
q_RunDO := iq_stPtm.q_RunDO;
q_xRemote := iq_stPtm.q_xRemote; // remote out
END_ACTION

ACTION ACT_Logger:
//STATE Logger
IF NOT i_xExtIlkOK AND ePrevState = pumpRUNNING THEN
         fbLogger(sMsg:='Lost external interlock while pump was running.', eSevr:=TcEventSeverity.Critical);
END_IF


IF ePrevState <> iq_stPTM.eState THEN
      CASE iq_stPTM.eState OF
        pumpFAULT:
            fbLogger(sMsg:='Pump Fault.', eSevr:=TcEventSeverity.Critical);
          pumpSTOPPED:
            fbLogger(sMsg:='Pump stopped.', eSevr:=TcEventSeverity.Critical);
        pumpSTARTING:
            fbLogger(sMsg:='Pump starting.', eSevr:=TcEventSeverity.Info);
        pumpRUNNING:
            fbLogger(sMsg:='Pump running.', eSevr:=TcEventSeverity.Info);
      END_CASE
      ePrevState := iq_stPTM.eState;
  END_IF

// ILK logger



// Log Action
tAction(CLK:=  iq_stPTM.q_RunDO);
IF tAction.Q THEN fbLogger(sMsg:='Pump commanded to start', eSevr:=TcEventSeverity.Info); END_IF


// Log FAULT
tFault(CLK:= NOT iq_stPTM.i_xFault);
IF tFault.Q THEN fbLogger(sMsg:='Pump Lost Alarm OK bit', eSevr:=TcEventSeverity.Critical); END_IF
END_ACTION

ACTION ACT_Persistent:
(*On first PLC pass, load the persistent value into the structrue variable*)
IF (SUPER^.bRestorePersistentData) THEN
    SUPER^.bRestorePersistentData	:= FALSE;
    IF (rBackingPressureSP <> 0) THEN
        iq_stPTM.rBackingPressureSP := rBackingPressureSP;
    END_IF;
    IF (rInletPressureSP <> 0) THEN
        iq_stPTM.rInletPressureSP := rInletPressureSP;
    END_IF;
END_IF
(*Check if a new value has been written in the structure variable copy it to the persistent variable*)
IF NOT (iq_stPTM.rBackingPressureSP = rBackingPressureSP) THEN
    rBackingPressureSP:= iq_stPTM.rBackingPressureSP;
END_IF;

IF NOT (iq_stPTM.rInletPressureSP = rInletPressureSP) THEN
    rInletPressureSP := iq_stPTM.rInletPressureSP;
END_IF;
END_ACTION

METHOD PUBLIC M_Run : BOOL
VAR_INPUT
    run:bool; // set to true to run, false to stop;
END_VAR

this^.iq_stPtm.xRunSW := run;
END_METHOD

END_FUNCTION_BLOCK

// ---- POUs/Functions/Pumps/FB_PTM_Pfeiffer.TcPOU
(* This function block does basic controls FOR the Pfeiffer Turbo pump connected to the TM700 and TC400 Controllers.
 Turns off pump in the event of errors/ warnings. Provides interlocking interface.*)
FUNCTION_BLOCK FB_PTM_Pfeiffer EXTENDS FB_Pump
VAR_INPUT
    i_xExtIlkOK : BOOL; // Connect to external interlock logic, TRUE if not used.
END_VAR
VAR_OUTPUT
    {attribute 'pytmc' := '
    pv:
    '}
    iq_stPTM : ST_PfeifferPTM;
END_VAR
VAR
    TOF_RESET: TON :=(PT:=T#1S);
    (*IO*)
    i_xAtSpd AT%I*: BOOL; // Normaml operation when true
    i_xFaultNC AT%I*: BOOL; // Error
    i_xWarn AT%I*: BOOL;
     i_xRemote AT%I*: BOOL;

    q_RunDO AT%Q*: BOOL; // Start/Stop for TC110 link this output to the Pumping station bit
    q_PumpingStation AT%Q*: BOOL; // Start/Stop interlock
    q_xRemote AT%Q*: BOOL;
    q_xReset AT%Q*: BOOL;
END_VAR

(* Basic pump supervisory section *)

q_xRemote := TRUE;
(* Interlock Sum *)
iq_stPtm.xExtRunOk:= i_xExtILKOk;
//For compatability with TC110
(*IF iq_stPTM.xExtRunOk THEN
    q_PumpingStation:= TRUE;
ELSE
    q_PumpingStation:= FALSE;
END_IF*)

IF iq_stPTM.xExtRunOk AND NOT (iq_stPTM.i_xFault) (*OR iq_stPTM.i_xTempFault)*) THEN
    iq_stPTM.q_RunDO:=iq_stPTM.xRunSW;
    q_PumpingStation:=iq_stPTM.xRunSW;
ELSE
    iq_stPTM.xRunSW:=FALSE;
    iq_stPTM.q_RunDO:=FALSE;
    q_PumpingStation:=FALSE;
END_IF


(*Pump STATE*)
IF iq_stPtm.i_xFault THEN
    iq_stPtm.eState := pumpFAULT;
ELSIF NOT iq_stPtm.q_RunDO AND NOT iq_stPTM.i_xFault THEN
    iq_stPtm.eState := pumpSTOPPED;
ELSIF NOT iq_stPtm.i_xAtSpd  AND iq_stPtm.q_RunDO THEN
    iq_stPtm.eState := pumpSTARTING;
ELSIF iq_stPtm.i_xAtSpd AND iq_stPtm.q_RunDO THEN
    iq_stPtm.eState := pumpRUNNING;
ELSE
    iq_stPtm.eState := pumpFAULT;
END_IF

(*Error Reset*)
(* to reset the Reset Bit *)
 IF (iq_stPTM.xResetSW ) THEN
    iq_stPTM.q_xReset := TRUE;
    q_PumpingStation := TRUE;
 END_IF

 IF (iq_stPTM.xResetSW) AND (iq_stPTM.i_xFault)  THEN
    q_PumpingStation := TRUE;
 END_IF
 TOF_RESET (IN:= iq_stPTM.q_xReset, Q => );
 IF TOF_RESET.Q THEN
    iq_stPTM.q_xReset:= FALSE;
    iq_stPTM.xResetSW := FALSE;
 END_IF

(*Soft IO Mapping*)
ACT_IO();
// Log States and triggers
ACT_Logger();
(*Load or save the persistent variables*)
ACT_Persistent();

ACTION ACT_IO:
(*outputs*)
q_RunDO := iq_stPTM.q_RunDO;
q_xReset := iq_stPTM.q_xReset;
//q_xRemote := iq_stPTM.
//q_PumpingStation AT%Q*: BOOL; // Start/Stop

(*inputs*)
iq_stPTM.i_xAtSpd:= i_xAtSpd;
iq_stPTM.i_xFault:= NOT i_xFaultNC;
iq_stPTM.i_xWarn:=  	i_xWarn ;
END_ACTION

ACTION ACT_Logger:
//STATE Logger
IF NOT i_xExtIlkOK AND ePrevState = pumpRUNNING THEN
         fbLogger(sMsg:='Lost external interlock while pump was running.', eSevr:=TcEventSeverity.Critical);
END_IF


IF ePrevState <> iq_stPTM.eState THEN
      CASE iq_stPTM.eState OF
        pumpFAULT:
            fbLogger(sMsg:='Pump Fault.', eSevr:=TcEventSeverity.Critical);
          pumpSTOPPED:
            fbLogger(sMsg:='Pump stopped.', eSevr:=TcEventSeverity.Critical);
        pumpSTARTING:
            fbLogger(sMsg:='Pump starting.', eSevr:=TcEventSeverity.Info);
        pumpRUNNING:
            fbLogger(sMsg:='Pump running.', eSevr:=TcEventSeverity.Info);
      END_CASE
      ePrevState := iq_stPTM.eState;
  END_IF

// ILK logger



// Log Action
tAction(CLK:=  iq_stPTM.q_RunDO);
IF tAction.Q THEN fbLogger(sMsg:='Pump commanded to start', eSevr:=TcEventSeverity.Info); END_IF


// Log FAULT
tFault(CLK:= NOT iq_stPTM.i_xFault);
IF tFault.Q THEN fbLogger(sMsg:='Pump Lost Alarm OK bit', eSevr:=TcEventSeverity.Critical); END_IF
END_ACTION

ACTION ACT_Persistent:
(*On first PLC pass, load the persistent value into the structrue variable*)
IF (SUPER^.bRestorePersistentData) THEN
    SUPER^.bRestorePersistentData	:= FALSE;
    IF (rBackingPressureSP <> 0) THEN
        iq_stPTM.rBackingPressureSP := rBackingPressureSP;
    END_IF;
    IF (rInletPressureSP <> 0) THEN
        iq_stPTM.rInletPressureSP := rInletPressureSP;
    END_IF;
END_IF
(*Check if a new value has been written in the structure variable copy it to the persistent variable*)
IF NOT (iq_stPTM.rBackingPressureSP = rBackingPressureSP) THEN
    rBackingPressureSP:= iq_stPTM.rBackingPressureSP;
END_IF;

IF NOT (iq_stPTM.rInletPressureSP = rInletPressureSP) THEN
    rInletPressureSP := iq_stPTM.rInletPressureSP;
END_IF;
END_ACTION

METHOD PUBLIC M_Run : BOOL
VAR_INPUT
    run:bool; // set to true to run, false to stop;
END_VAR

this^.iq_stPtm.xRunSW := run;
END_METHOD

METHOD PUBLIC M_Serial_IO : BOOL
VAR_INPUT
    st_Pfeiffer_RBK: ST_PfeifferStatus;
END_VAR
VAR_IN_OUT
    st_Pfeiffer_CTRL: ST_PfeifferControl;
END_VAR
(* This function block is used to map the IO points from the pfeiffer structures
to the generic turbo structures *)
(*
if (bInit) Then
    bInit := False;
    st_Pfeiffer_CTRL.diSetRotationSpeed_309 := st_Pfeiffer_RBK.diActiveRotationSpeed_309;
END_IF*)

(* Controls *) (* Controls is via DIO*)
//st_Pfeiffer_CTRL.xPumpingStation_010 := iq_stPTM.q_RunDO;
//st_Pfeiffer_CTRL.xMotorPump_023 := 1; //Setting always true because parameter 10 alone can enable/disable the pump
//st_Pfeiffer_CTRL.uiPowerPct_708 := iq_stPTM.q_uiPowerPct;
//st_Pfeiffer_CTRL.xErrorAck_009 := iq_stPTM.xResetSW;



(* Readbacks *)
iq_stPTM.i_xAccel := st_Pfeiffer_RBK.xPumpAccelerating_307;
//iq_stPTM.i_xAtSpd := st_Pfeiffer_RBK.xRotationSpeedAttn_306; The Atspd is already linked via Digital I/Os
iq_stPTM.i_diCurSpd := st_Pfeiffer_RBK.diActiveRotationSpeed_309;
iq_stPTM.i_diPwr := st_Pfeiffer_RBK.diDrivePower_316;
iq_stPTM.i_diElecTemp := st_Pfeiffer_RBK.diTempElec_326;
iq_stPTM.i_diBtmTemp := st_Pfeiffer_RBK.diTempPmpBot_330;
iq_stPTM.i_diBrngTemp := st_Pfeiffer_RBK.diTempBearng_342;
iq_stPTM.i_diMtrTemp := st_Pfeiffer_RBK.diTempMotor_346;
iq_stPTM.i_uiPowerPctRbk := st_Pfeiffer_RBK.uiPowerPct_708;
iq_stPTM.i_rCurrentMon :=  LREAL_TO_REAL(st_Pfeiffer_RBK.lrDriveCurrent_310);
iq_stPTM.xCommTimeout	:=	st_Pfeiffer_RBK.xTimeout;
iq_stPTM.i_iErrorCode := st_Pfeiffer_RBK.iErrorCode_303;
iq_stPTM.i_iWarningCode := st_Pfeiffer_RBK.iWarningCode_303;

(* Check that error acknowledgment is processed *)
IF st_Pfeiffer_RBK.xErrorAcknowledged THEN
    st_Pfeiffer_RBK.xErrorAcknowledged := FALSE;
    st_Pfeiffer_CTRL.xErrorAck_009 := FALSE;
    iq_stPTM.xResetSW := FALSE;
END_IF

IF st_Pfeiffer_RBK.sErrorCode_303 = '' THEN
    ;
ELSIF st_Pfeiffer_RBK.iErrorCode_303 <> 0 THEN
iq_stPTM.i_xFault := TRUE;
ELSE
iq_stPTM.i_xFault := FALSE;
END_IF

st_Pfeiffer_CTRL.xSetSpdMode_026:= iq_stPTM.q_bSetSpd;
iq_stPTM.i_dSetSpd := LIMIT (0, iq_stPTM.i_dSetSpd, 1500); // 1500 nominal frequency
IF ( iq_stPTM.i_dSetSpd <>0) THEN
    st_Pfeiffer_CTRL.iSetRotationSpeed_707 := DINT_TO_INT(iq_stPTM.i_dSetSpd * 100/1500);
    st_Pfeiffer_CTRL.iSetRotationSpeed_707 := LIMIT(20, st_Pfeiffer_CTRL.iSetRotationSpeed_707 ,100); // Manual Page 18
END_IF
END_METHOD

METHOD PUBLIC M_SetBackingSP
VAR_INPUT
    i_fBackingPressureSP : REAL;
END_VAR
iq_stPTM.rBackingPressureSP := i_fBackingPressureSP;
END_METHOD

METHOD PUBLIC M_SetForelineSP
VAR_INPUT
    i_fForelinePressureSP : REAL;
END_VAR
iq_stPTM.rForelineSP := i_fForelinePressureSP;
END_METHOD

END_FUNCTION_BLOCK

// ---- POUs/Functions/Pumps/FB_PTM_TurboDrive.TcPOU
(* This Function block provides basic turbo control for Leybold Turbo Drive 300, Turbo Drive 400 *)
(* TD20 Classic Via Remote X1 Connector 9-way PLC interface*)
(* When serial interface is implemented, call Method M_Serial_IO after fb instantiation, in order to add the serial status *)
FUNCTION_BLOCK FB_PTM_TurboDrive EXTENDS FB_Pump
VAR_INPUT
    i_xExtILKOk : BOOL; // Connect to external interlock logic, TRUE if not used.
END_VAR
VAR_OUTPUT
    {attribute 'pytmc' := '
    pv:
    '}
    iq_stPtm	:	ST_LeyboldPTM;
END_VAR
VAR

    xRunOk	:	BOOL;
    tofRemoteDelay	:	TOF;


    (*IO*)
    i_xAtSpd AT%I*: BOOL; // Normaml operation when true
    i_xFaultNC AT%I*: BOOL; // Error Active when no Error is present
    q_RunDO AT%Q*: BOOL; // Start/Stop
END_VAR

(* Basic Turbo Control *)
(* This Function block provides basic turbo control for Leybold Turbo Drive 300, Turbo Drive 400 *)
(* TD20 Classic Via Remote X1 Connector 9-way PLC interface*)
(* M. Ghaly Jan. 2019 *)

(* Interlock Sum *)
iq_stPtm.xExtRunOk:= i_xExtILKOk;
xRunOk := iq_stPtm.xExtRunOk AND iq_stPtm.i_xNCError;

(* Basic pump supervisory section *)
IF xRunOk THEN
    q_RunDO := iq_stPTM.xRunSW;
ELSE
    iq_stPtm.xRunSW:=FALSE;
    q_RunDO:=FALSE;
END_IF

(*Pump States*)
IF (iq_stPtm.i_xFault) THEN
        iq_stPtm.eState := pumpFAULT;
        iq_stPtm.xRunSW:=FALSE;
        q_RunDO:=FALSE;
ELSIF (iq_stPtm.q_RunDO) AND (iq_stPtm.i_xAtSpd) THEN
        iq_stPtm.eState := pumpRUNNING;
ELSIF (iq_stPtm.q_RunDO) AND NOT (iq_stPtm.i_xAtSpd) THEN
        iq_stPtm.eState := pumpSTARTING;
ELSIF NOT (iq_stPtm.q_RunDO) THEN
        iq_stPtm.eState := pumpSTOPPED;
ELSE
    iq_stPtm.eState := pumpFAULT;
END_IF;


(*I/O soft mapping*)
ACT_IO();
// Log States and triggers
This^.ACT_Logger();
(*Load or save the persistent variables*)
ACT_Persistent();

ACTION ACT_IO:
(*Inputs*)
iq_stPtm.i_xAtSpd := i_xAtSpd;
iq_stPtm.i_xNCError := i_xFaultNC;
iq_stPtm.i_xFault := NOT i_xFaultNC;



(*Outputs*)
iq_stPtm.q_RunDO := q_RunDO;
END_ACTION

ACTION ACT_Logger:
//STATE Logger
// ILK logger
IF NOT i_xExtIlkOK AND ePrevState = pumpRUNNING THEN
         fbLogger(sMsg:='Lost external interlock while pump was running.', eSevr:=TcEventSeverity.Critical);
END_IF


IF ePrevState <> iq_stPTM.eState THEN
      CASE iq_stPTM.eState OF
        pumpFAULT:
            fbLogger(sMsg:='Pump Fault.', eSevr:=TcEventSeverity.Critical);
          pumpSTOPPED:
            fbLogger(sMsg:='Pump stopped.', eSevr:=TcEventSeverity.Critical);
        pumpSTARTING:
            fbLogger(sMsg:='Pump starting.', eSevr:=TcEventSeverity.Info);
        pumpRUNNING:
            fbLogger(sMsg:='Pump running.', eSevr:=TcEventSeverity.Info);
      END_CASE
      ePrevState := iq_stPTM.eState;
  END_IF

// Log Action
tAction(CLK:=  iq_stPTM.q_RunDO);
IF tAction.Q THEN fbLogger(sMsg:='Pump commanded to start', eSevr:=TcEventSeverity.Info); END_IF


// Log FAULT
tFault(CLK:= NOT iq_stPTM.i_xFault);
IF tFault.Q THEN fbLogger(sMsg:='Pump Lost Alarm OK bit', eSevr:=TcEventSeverity.Critical); END_IF
END_ACTION

ACTION ACT_Persistent:
(*On first PLC pass, load the persistent value into the structrue variable*)
IF (SUPER^.bRestorePersistentData) THEN
    SUPER^.bRestorePersistentData	:= FALSE;
    IF (rBackingPressureSP <> 0) THEN
        iq_stPTM.rBackingPressureSP := rBackingPressureSP;
    END_IF;
    IF (rInletPressureSP <> 0) THEN
        iq_stPTM.rInletPressureSP := rInletPressureSP;
    END_IF;
END_IF
(*Check if a new value has been written in the structure variable copy it to the persistent variable*)
IF NOT (iq_stPTM.rBackingPressureSP = rBackingPressureSP) THEN
    rBackingPressureSP:= iq_stPTM.rBackingPressureSP;
END_IF;

IF NOT (iq_stPTM.rInletPressureSP = rInletPressureSP) THEN
    rInletPressureSP := iq_stPTM.rInletPressureSP;
END_IF;
END_ACTION

METHOD PUBLIC M_Run : BOOL
VAR_INPUT
    run:bool; // set to true to run, false to stop;
END_VAR

this^.iq_stPtm.xRunSW := run;
END_METHOD

METHOD PUBLIC M_Serial_IO : BOOL
VAR_INPUT
    i_st_TD20_RBK			: ST_TD20Status;
END_VAR

(* This function block is used to map the IO points from the Oerlikon structures
to the generic turbo structures *)

(* Readbacks *)
iq_stPTM.i_xAccel := i_st_TD20_RBK.wStatusWord.4;
iq_stPTM.i_xDecel := i_st_TD20_RBK.wStatusWord.5;
//iq_stPTM.i_xAtSpd := i_st_TD20_RBK.wStatusWord.10;
iq_stPTM.i_xRemote := i_st_TD20_RBK.wStatusWord.15; (* Remote control enabled *)
iq_stPTM.i_diCurSpd := WORD_TO_DINT(i_st_TD20_RBK.wFrequency_P3);
iq_stPTM.i_rCurrentMon := WORD_TO_INT(i_st_TD20_RBK.wMotorCurrent_P5)*0.1; (*Current in units 0.1 A, TD20 manual page 23*)
iq_stPTM.i_diPwr := LREAL_TO_DINT(WORD_TO_DINT(i_st_TD20_RBK.wMotorCurrent_P5 * i_st_TD20_RBK.wVoltage_P4)*0.01); (*Current in units 0.1 A and voltage in units 0.1V, TD20 manual page 23*)
iq_stPTM.i_diElecTemp := WORD_TO_DINT(i_st_TD20_RBK.wConverterTemp_P11);
iq_stPTM.i_rTempMon := WORD_TO_INT(i_st_TD20_RBK.wPumpTemp_P127);

(* Faults and warnings *)
//iq_stPTM.i_xFault := i_st_TD20_RBK.wStatusWord.3;
iq_stPTM.i_xTempFault := i_st_TD20_RBK.wStatusWord.7; (* specified as a temperature warning but it could be a fault *)
iq_stPTM.i_xWarn := i_st_TD20_RBK.wStatusWord.14; (* warning summary bit *)
END_METHOD

METHOD PUBLIC M_SetBackingSP
VAR_INPUT
    i_fBackingPressureSP : REAL;
END_VAR
iq_stPtm.rBackingPressureSP := i_fBackingPressureSP;
END_METHOD

METHOD PUBLIC M_SetForelineSP
VAR_INPUT
    i_fForelinePressureSP : REAL;
END_VAR
iq_stPtm.rForelineSP := i_fForelinePressureSP;
END_METHOD

END_FUNCTION_BLOCK

// ---- POUs/Functions/Pumps/FB_ScrollPump.TcPOU
(* This Function block provides basic  control for Scroll Pumps *)
(* Turn on scroll pump if the Turbo Vent Valve is closed. *)
(* Cannot turn off scroll pump if turb is running. delay scroll off 150s.*)

FUNCTION_BLOCK FB_ScrollPump
VAR_IN_OUT

END_VAR
VAR_OUTPUT
    {attribute 'pytmc' := '
    pv:
    '}
    iq_stPFO	:	ST_RoughPump;
END_VAR
VAR_INPUT
    TurboIsON : BOOL;
    xExtIlk : BOOL;
END_VAR
VAR
    Tmr_TOF : TOF;
    tTimerDuration : Time:= T#150S;
    //Previous_RunSW : BOOL;
    // Digital Output to be linked
    q_xRunDo AT%Q*	:   BOOL;
END_VAR

//Turn on scroll pump if the Turbo Vent Valve is closed. So you are not just
// pumping air and accomplishing nothing

// cannot turn off scroll pump if turb is running. delay scroll off 150s.
iq_stPFO.xIlkOK := xExtIlk;// and NOT Tmr_TOF.Q;

Tmr_TOF(IN:=TurboIsON, PT := tTimerDuration);

IF iq_stPFO.xIlkOK THEN
    iq_stPFO.q_xRunDo := (Tmr_TOF.Q OR iq_stPFO.pv_xRunSW);
ELSE
    iq_stPFO.q_xRunDo := FALSE;
END_IF

iq_stPFO.pv_xRunSW := iq_stPFO.q_xRunDo;

(*State evaluation*)
IF NOT iq_stPFO.q_xRunDo THEN
    iq_stPFO.eState := pumpSTOPPED;
ELSE
    iq_stPFO.eState := pumpRUNNING;
END_IF

(*soft io Mapping*)
IO();

ACTION IO:
q_xRunDo:= iq_stPFO.q_xRunDo;
END_ACTION

METHOD PUBLIC M_Run : BOOL
VAR_INPUT
    run:bool; // set to true to run, false to stop;
END_VAR

this^.iq_stPFO.pv_xRunSW := run;
END_METHOD

END_FUNCTION_BLOCK

// ---- POUs/Functions/Pumps/functions/FB_TurboExtLogic.TcPOU
(*deprecated*)
FUNCTION_BLOCK FB_TurboExtLogic
VAR_IN_OUT
    Turbo		:	ST_AgilentPTM;
END_VAR
VAR_INPUT
    BackingGauge:	ST_VG;
    InletGauge	:	ST_VG;
    VentValve	:	ST_VCC_NO;
    ScrollPump	:	ST_RoughPump;
END_VAR
VAR_OUTPUT
END_VAR
VAR
END_VAR

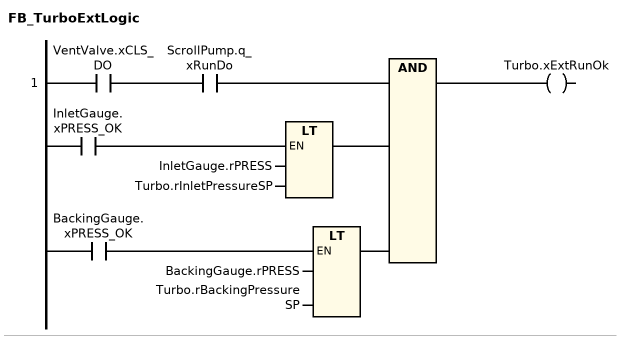
// NETWORK 1
Turbo.xExtRunOk := (VentValve.xCLS_DO AND ScrollPump.q_xRunDo) AND (InletGauge.xPRESS_OK AND InletGauge.rPRESS < Turbo.rInletPressureSP) AND (BackingGauge.xPRESS_OK AND BackingGauge.rPRESS < Turbo.rBackingPressureSP);

END_FUNCTION_BLOCK

// ---- POUs/Functions/Pumps/functions/F_TurboExtILK_NO.TcPOU
(* This function Block interfaces with a NO turbo valve*)
(* Mainly used in the FEE HXR GATT*)
FUNCTION F_TurboExtILK_NO : BOOL
VAR_INPUT
    Turbo		:	ST_PTM;
    BackingGauge:	ST_VG;
    InletGauge	:	ST_VG;
    VentValve	:	ST_VCC_NO; //NO type turbo valve
    ScrollPump	:	ST_RoughPump;
END_VAR

VAR
END_VAR

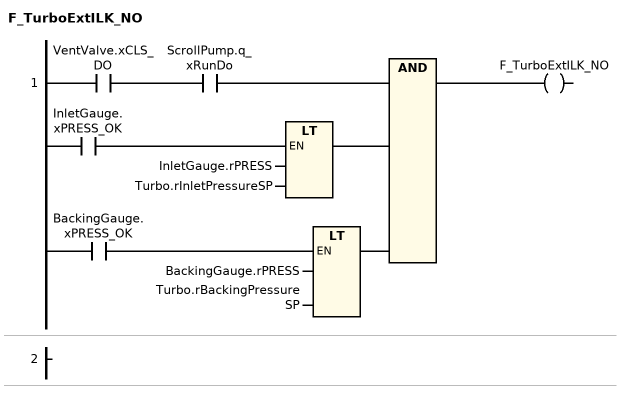
// NETWORK 1
F_TurboExtILK_NO := (VentValve.xCLS_DO AND ScrollPump.q_xRunDo) AND (InletGauge.xPRESS_OK AND InletGauge.rPRESS < Turbo.rInletPressureSP) AND (BackingGauge.xPRESS_OK AND BackingGauge.rPRESS < Turbo.rBackingPressureSP);

// NETWORK 2

END_FUNCTION

// ---- POUs/Functions/Pumps/functions/F_TurboExtILKLogic.TcPOU

(* This function evaluates the Turbo ILK logic*)
(* The Turbo shall not Run if the vent valve is open*)
(* The function also switches off the Turbo if the Inlet pressure or the backing Pressure*)
(* are higher than the configured set point*)
FUNCTION F_TurboExtILKLogic : BOOL
VAR_INPUT
    Turbo		:	ST_PTM;
    BackingGauge:	ST_VG;
    InletGauge	:	ST_VG;
    VentValve	:	ST_VVC;
    ScrollPump	:	ST_RoughPump;
END_VAR

VAR
END_VAR

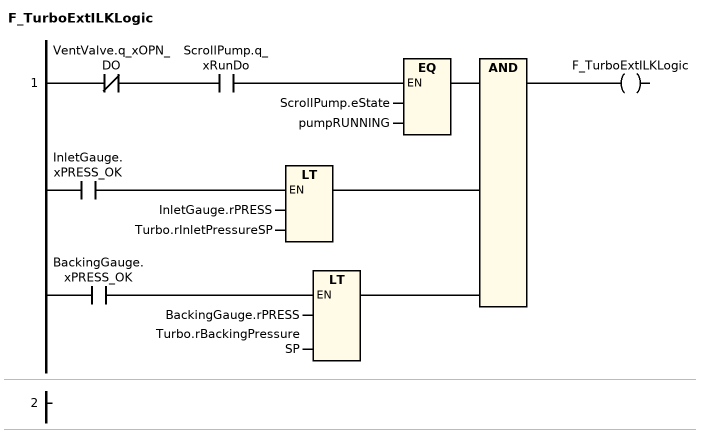
// NETWORK 1
F_TurboExtILKLogic := (NOT VentValve.q_xOPN_DO AND ScrollPump.q_xRunDo AND ScrollPump.eState = pumpRUNNING) AND (InletGauge.xPRESS_OK AND InletGauge.rPRESS < Turbo.rInletPressureSP) AND (BackingGauge.xPRESS_OK AND BackingGauge.rPRESS < Turbo.rBackingPressureSP);

// NETWORK 2

END_FUNCTION

// ---- POUs/Functions/Pumps/functions/F_TurboExtILKLogic_2.TcPOU

(* This function evaluates the Turbo ILK logic*)
(* The function switches off the Turbo if the Inlet pressure or the backing Pressure*)
(* are higher than the configured set point*)
FUNCTION F_TurboExtILKLogic_2 : BOOL
VAR_INPUT
    Turbo		:	ST_PTM;
    BackingGauge:	ST_VG;
    InletGauge	:	ST_VG;
    ScrollPump	:	ST_RoughPump;
END_VAR
VAR
END_VAR

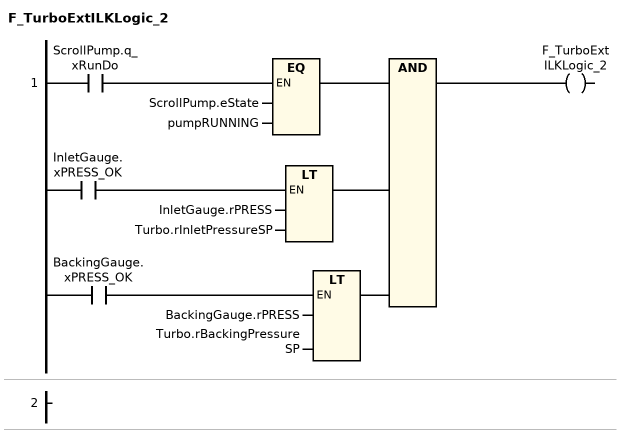
// NETWORK 1
F_TurboExtILKLogic_2 := (ScrollPump.q_xRunDo AND ScrollPump.eState = pumpRUNNING) AND (InletGauge.xPRESS_OK AND InletGauge.rPRESS < Turbo.rInletPressureSP) AND (BackingGauge.xPRESS_OK AND BackingGauge.rPRESS < Turbo.rBackingPressureSP);

// NETWORK 2

END_FUNCTION

// ---- POUs/Functions/Pumps/functions/F_TurboExtILK_NO_1.TcPOU
(* This function Block interfaces with a NO turbo valve*)
(* Mainly used in the FEE HXR GATT*)
FUNCTION F_TurboExtILK_NO_1 : BOOL
VAR_INPUT
    Turbo		:	ST_PTM;
    BackingGauge:	ST_VG;
    InletGauge	:	ST_VG;
    VentValve	:	ST_VCC_NO; //NO type turbo valve
    ScrollPump	:	ST_RoughPump;
END_VAR

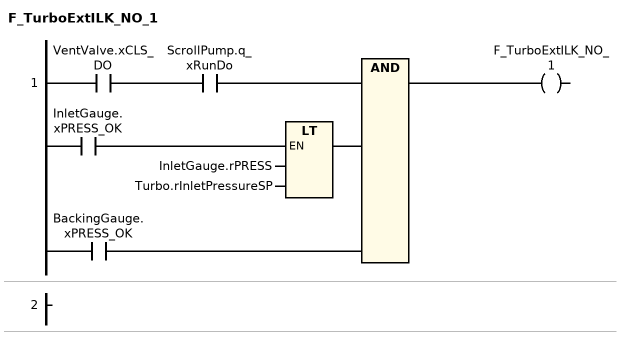
// NETWORK 1
F_TurboExtILK_NO_1 := (VentValve.xCLS_DO AND ScrollPump.q_xRunDo) AND (InletGauge.xPRESS_OK AND InletGauge.rPRESS < Turbo.rInletPressureSP) AND BackingGauge.xPRESS_OK;

// NETWORK 2

END_FUNCTION

// ---- POUs/Functions/Pumps/Interfaces/FB_PIP_Interface_In.TcPOU
(* This function block is created for interface devices between different PLC*)
(* Not all the Variables in the original structure is required, just few signals *)
(* They have to be linked to the custom created variables on the EL6692/5 primary side*)
FUNCTION_BLOCK FB_PIP_Interface_In
VAR_INPUT
END_VAR
VAR_OUTPUT
    VG : ST_VG;
END_VAR
VAR
    i_rPRESS AT%I*: REAL;  //This is the human-readable pressure
    i_xAT_VAC AT%I*: BOOL;
    i_xPRESS_OK AT%I*: BOOL;
    i_xIs_Connected AT%I*: BOOL;
END_VAR

(* This function block is created for interface devices between different PLC*)
(* Not all the Variables in the original structure is required, just few signals *)
(* They have to be linked to the custom created variables on the EL6692/5 primary side*)

VG.rPRESS := i_rPRESS;
VG.xAT_VAC := i_xAT_VAC;
VG.xPRESS_OK := i_xPRESS_OK;


IF NOT(i_xIs_Connected) THEN
    i_xPRESS_OK := FALSE;
END_IF

END_FUNCTION_BLOCK

// ---- POUs/Functions/Pumps/Interfaces/FB_PIP_Interface_Out.TcPOU
(* This function block is created for interface devices between different PLC*)
(* Not all the Variables in the original structure is required, just few signals *)
(* They have to be linked to the custom created variables on the EL6692/5 primary side*)
FUNCTION_BLOCK FB_PIP_Interface_Out
VAR_INPUT
    VG : ST_VG;
END_VAR
VAR_OUTPUT
END_VAR
VAR
    i_rPRESS AT%Q*: REAL;
    i_xAT_VAC AT%Q*: BOOL;
    i_xPRESS_OK AT%Q*: BOOL;
END_VAR

(* This function block is created for interface devices between different PLC*)
(* Not all the Variables in the original structure is required, just few signals *)
(* They have to be linked to the custom created variables on the EL6692/5 primary side*)

i_rPRESS:=VG.rPRESS;
i_xAT_VAC:= VG.xAT_VAC;
i_xPRESS_OK:=VG.xPRESS_OK;

END_FUNCTION_BLOCK

// ---- POUs/Functions/Pumps/Interfaces/FB_TPIP_ADS.TcPOU
(* This function block is created for interface devices between different PLC*)
(* Not all the Variables in the original structure is required, just few signals *)
(* The variable values are read via ADS using the symbol name*)
FUNCTION_BLOCK FB_TPIP_ADS Extends FB_ADS
VAR_INPUT
    sNetId : String; //NetID of the Destination PLC controller
    nPort : uint; // port number
    sVarName : string;// the variable name of the declared pip/pin function block.
    iWatchdog:UDINT;//The watchdog variable name written to by the remote plc
END_VAR
VAR_OUTPUT
    {attribute 'pytmc' := 'pv:'}
    IG : ST_VG;
    bError: BOOL;
END_VAR
VAR
    fb_CheckWatchdog: FB_CheckWatchdog;
    fb_Read_VG: FB_ReadAdsSymByName;
    ftReset: F_TRIG;
    xFirstPass: BOOL:= true;

END_VAR


ftReset(CLK:= fb_Read_VG.bBusy OR xFirstPass);
xFirstPass := false;
(*calling ADS read function*)

fb_Read_VG(
    bRead:=ftReset.Q ,
    sNetId:= sNetId,
    nPort:= nPort,
    sVarName:= CONCAT(sVarName,'.q_IG'),
    nDestAddr:= ADR(IG),
    nLen:= SIZEOF(IG),
    tTimeout:= ,
    eComMode:=eAdsComModeFastCom ,
    bBusy=> ,
    bError=> ,
    nErrorId=> );


(*Error*)
fb_CheckWatchdog(
    bEnable:= TRUE,
    tWatchdogTime:= T#900ms,
    nCnt:= iWatchdog ,
    bWatchdog=> ,
    nLastCnt=> );

bError:= fb_Read_VG.bError OR fb_CheckWatchdog.bWatchdog;
tErrorPresent(CLK:=bError);

IF (fb_Read_VG.bError OR fb_CheckWatchdog.bWatchdog) THEN
IG.xPRESS_OK := FALSE;
END_IF;

(*Logger*)
ACT_Logger();

ACTION ACT_Logger:
IF tErrorPresent.Q THEN
 IF(fb_Read_VG.bError) THEN fbLogger(sMsg:='ADS Read Error', eSevr:=TcEventSeverity.Critical); END_IF;
 IF(fb_CheckWatchdog.bWatchdog) THEN fbLogger(sMsg:='ADS Watchdog Error', eSevr:=TcEventSeverity.Critical); END_IF;
END_IF
END_ACTION

END_FUNCTION_BLOCK

// ---- POUs/Functions/Valves/FB_Kashiyama_VRC.TcPOU
(* Main Kashiyama gate valve permit to be open when:
        1. pump is NORMAL operating status, and
        2. chamber pressure is below HighSP or pump is at LowSpeed state.
    it will close if chamber pressure is below than lowSP for 180s.
*)
FUNCTION_BLOCK FB_Kashiyama_VRC
VAR_IN_OUT

END_VAR
VAR_OUTPUT
    {attribute 'pytmc' := ' pv:'}
    q_stValve : ST_VRC;
END_VAR
VAR_INPUT
    Pump : ST_KashiyamaDryPump;//Kashyiama pump
    i_xExtILK_OK : BOOL; //Connect to Interlock logic condition(e.g F_TURBO_VRC_ILK Function), otherwise, Set to True if the valve is not interlocked
    Gauge : ST_VG;// Pressure Gauge
    i_xOverrideMode : BOOL;
END_VAR
VAR
    At_HiVac : BOOL;
    tmrTP : TP;
    tmrPT: TIME := T#180S;
    v1: BOOL;
    tonOvrd	:	TON;
    tonDelOK : TON;
    rtOK	:	R_TRIG;

    (*IO*)
    i_xOpnLS	AT%I*: BOOL;
    i_xClsLS	AT%I*: BOOL;
    q_xOPN_DO	AT%Q*: BOOL;

END_VAR

(* Main Kashiyama gate valve permit to be open when:
        1. pump is NORMAL operating status, and
        2. chamber pressure is below HighSP or pump is at LowSpeed state.
    it will close if chamber pressure is below than lowSP for 60s.
*)
(*
      For main Kayshiyama pump's gate valve:
        Pump LowSP is MU100 base pressure (20 mTorr)
        Pump HighSP is 600 Torr;
      Second Kayshiyama pump allow Gas Attenuator operating at higher pressure,
      it's gate valve is to be open when Gas Attenuator chamber pressure is above lowSP.
*)


///Check valve postion
IF NOT q_stValve.i_xClsLS AND q_stValve.i_xOpnLS THEN
    q_stValve.eState:=OPEN;
ELSIF q_stValve.i_xClsLS AND NOT q_stValve.i_xOpnLS THEN
    q_stValve.eState:=CLOSED;
ELSIF NOT q_stValve.i_xClsLS AND NOT q_stValve.i_xOpnLS THEN
    q_stValve.eState:=MOVING;
ELSE
    q_stValve.eState:=INVALID;
END_IF

//valve open interlock
q_stValve.xOPN_OK := Pump.i_xIsRun AND Pump.RdyTmr <= 0.0 AND (Gauge.rPRESS < Pump.HighSP OR Pump.q_xLspdDo) AND i_xExtILK_OK;


(* Override logic *)
(* Goal: give ability to override, but do so in a way that people won't forget it.
Solution: Override only after ten seconds of override, protect against blips,
when the valve permission goes true for more than ten seconds consistently, remove override
*)

tonDelOK(IN:=q_stValve.xOPN_OK, PT:=T#10S);
rtOK(CLK:=tonDelOK.Q);
IF rtOK.Q THEN q_stValve.pv_xOvrdOpn :=FALSE; END_IF

//Override timer
tonOvrd(IN:=q_stValve.pv_xOvrdOpn, PT:=T#10S);


(* Here's where the valve closes *)
IF NOT q_stValve.xOPN_OK AND NOT tonOvrd.Q THEN
q_stValve.pv_xOPN_SW := FALSE;
END_IF

At_HiVac := Gauge.xPRESS_OK AND Gauge.rPRESS < Pump.LowSP;
tmrTP (IN := At_HiVac AND q_stValve.q_xOPN_DO , PT := tmrPT);

IF At_HiVac AND q_stValve.q_xOPN_DO AND NOT tmrTP.Q THEN
    q_stValve.pv_xOPN_SW := FALSE ;
END_IF

(* Here's where the valve opens *)
q_stValve.q_xOPN_DO := (q_stValve.pv_xOPN_SW AND q_stValve.xOPN_OK) OR (tonOvrd.Q AND i_xOverrideMode);

(*Soft IO Mapping*)
ACT_IO();

ACTION ACT_IO:
(*inputs*)
q_stValve.i_xOpnLS := 	i_xOpnLS;
q_stValve.i_xClsLS:=	i_xClsLS;
(*outputs*)
q_xOPN_DO:= q_stValve.q_xOPN_DO;
END_ACTION

END_FUNCTION_BLOCK

// ---- POUs/Functions/Valves/FB_MKS248.TcPOU
(* MKS248 valve using MKS1249 Drive Module *)
FUNCTION_BLOCK FB_MKS248
VAR_INPUT
    i_xExtIlkOK	:	BOOL; //External Interlock, SET to TRUE if not used
    i_rReqPos	:	REAL; //Requested position
END_VAR
VAR_OUTPUT
    {attribute 'pytmc' := 'pv:'}
    iq_stVFN	:	ST_VCN; //Needle valve structure
END_VAR
VAR CONSTANT
    rOpenVoltage	:	REAL := 9.8;
    rCloseVoltage	:	REAL := 0;
END_VAR
VAR
    // Requested voltage
    rReqVoltage: REAL := 0;
    (*IO*)
    q_iRawPosition AT%Q* :INT;
END_VAR

(* MKS248 valve using MKS1249 Drive Module *)


// Interlocking
iq_stVFN.xIlkOK := i_xExtIlkOK;
(*Checking which Control mode is selected*)
IF iq_stVFN.xIlkOK THEN
    IF iq_stVFN.eValveControl = OpenValve THEN
        iq_stVFN.rReqPosition := iq_stVFN.rUpperLimit;(*Percentage*)// iq_stVCN.rUpperLimit;
    ELSIF iq_stVFN.eValveControl = CloseValve THEN
        iq_stVFN.rReqPosition := 0; (*Percentage*)
    ELSIF iq_stVFN.eValveControl = ManualControl THEN
        iq_stVFN.rReqPosition := LIMIT(0, iq_stVFN.rReqPosition, iq_stVFN.rUpperLimit);
    ELSIF iq_stVFN.eValveControl = PressureControl THEN
        iq_stVFN.rReqPosition := LIMIT(0, i_rReqPos, iq_stVFN.rUpperLimit);
    END_IF
ELSE
    iq_stVFN.rReqPosition := 0;
    iq_stVFN.eValveControl := CloseValve;
END_IF

// Requested Voltage calculation
rReqVoltage := iq_stVFN.rReqPosition * (rOpenVoltage-rCloseVoltage)/100 + rCloseVoltage;
rReqVoltage := LIMIT(rCloseVoltage, rReqVoltage, rOpenVoltage); //The requested voltage should remain within this range
//Raw position calc
iq_stVFN.q_iRawPosition := REAL_TO_INT( 32767/10 * rReqVoltage);
(*IO Mapping*)
ACT_IO();

ACTION ACT_IO:
(*outputs*)
q_iRawPosition := iq_stVFN.q_iRawPosition;
END_ACTION

METHOD PUBLIC M_SetControlMode
VAR_INPUT
    i_eValveControlMode	:	E_VCN;
END_VAR
iq_stVFN.eValveControl := i_eValveControlMode;
END_METHOD

METHOD PUBLIC M_SetReqPosition
VAR_INPUT
    i_fReqPosition : REAL;
END_VAR
iq_stVFN.rReqPosition := i_fReqPosition;
END_METHOD

END_FUNCTION_BLOCK

// ---- POUs/Functions/Valves/FB_TurbVentvalve_NO.TcPOU
(* This function block impelemets Interlock for Agilent Turbo Vent Valve Normally Open*)
FUNCTION_BLOCK FB_TurbVentvalve_NO
VAR_OUTPUT
    {attribute 'pytmc' :=' pv:'}
    q_stValve : ST_VCC_NO;
END_VAR
VAR_INPUT
    i_stPTM	: ST_AgilentPTM; //Agilent Turbo Pump
END_VAR
VAR
    tofTmr 		: 	TOF;

    (*Output*)
    q_xCLS_DO AT%Q* : BOOL;
END_VAR

(*If the turbo is on, you cannot open the valve. In order to open the valve, you have to allow the turbopump
 to have already been turned off for 2 minutes and you have to press the open button on the vent valve

If the code looks confusing please use a truth table to verify*)

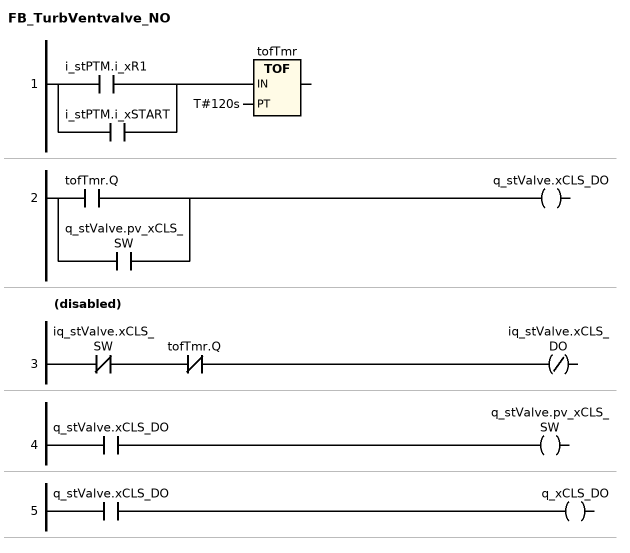
// NETWORK 1
tofTmr(IN := i_stPTM.i_xR1 OR i_stPTM.i_xSTART, PT := T#120s); // TOF

// NETWORK 2
q_stValve.xCLS_DO := tofTmr.Q OR q_stValve.pv_xCLS_SW;

// NETWORK 3 (disabled)
// iq_stValve.xCLS_DO := NOT (NOT iq_stValve.xCLS_SW AND NOT tofTmr.Q);

// NETWORK 4
q_stValve.pv_xCLS_SW := q_stValve.xCLS_DO;

// NETWORK 5
q_xCLS_DO := q_stValve.xCLS_DO;

ACTION ACT_IO:
(*outputs*)
q_xCLS_DO:= q_stValve.xCLS_DO;
END_ACTION

METHOD M_Close : BOOL
VAR_INPUT
        close:BOOL; //True to CLose, False to OPEN
END_VAR
This^.q_stValve.pv_xCLS_SW :=Close;
END_METHOD

END_FUNCTION_BLOCK

// ---- POUs/Functions/Valves/FB_VCN_VAT590.TcPOU
(* This function implements the Basic functions for the VAT590 needle valve*)
FUNCTION_BLOCK FB_VCN_VAT590 EXTENDS FB_Valve
VAR_INPUT
    bExtIlkOK : BOOL;        // External Interlock, SET to TRUE if not used
    IG : ST_VG;              // Input from a cold cathode gauge used in control loop
END_VAR
VAR_OUTPUT
    {attribute 'pytmc' := '
    pv:
    '}
    stVcnVat590	: ST_VCN_VAT590;       // Needle valve VAT590 structure
END_VAR
VAR CONSTANT
    cOpenPosition : REAL := 1E+5;      // Default position setpoint upper scale value
    cClosePosition : REAL := 0.0;      // Default position setpoint lower scale value
    cPresSPUpLim : REAL := 1E+6;       // Default pressure setpoint upper scale value
    cPresSPLowLim : REAL := 0;         // Default pressure setpoint lower scale value
    cMinPress : REAL := 1e-11;         // Default Min. pressure in Torr that can be used and requested
    cMaxPress : REAL := 1e-2;          // Default Max. pressure in Torr that can be used and requested
    cBasePress : REAL := 1E-11;        // Pressure sensor base value
    cPressRawSlope : REAL := 1E+5;     // Slope (in Units per decade) used for conversion of pressure in Torr to valve External Digital pressure sensor 1 input raw value (0-1000000)
    cPressRawBase : REAL := 1E+5;      // Valve analog output base(in Units per decade) defined for how much the curve is shifted

    cPressCtrl : ST_CoEIndSub := (nIndex := 16#2199, nSubIndex := 0); // Selected pressure controller CoE register
    cSensorDelay_AD : ST_CoEIndSub := (nIndex := 16#219A, nSubIndex := 0); // Adaptive DS controller Sensor Delay CoE register
    cRampTime_AD : ST_CoEIndSub := (nIndex := 16#219B, nSubIndex := 0); // Adaptive DS controller Ramp Time CoE register
    cRampMode_AD : ST_CoEIndSub := (nIndex := 16#219C, nSubIndex := 0); // Adaptive DS controller Ramp Mode CoE register
    cGainFactor_AD : ST_CoEIndSub := (nIndex := 16#219E, nSubIndex := 0); // Adaptive DS controller Gain factor CoE register
    cRampTime_FIX1 : ST_CoEIndSub := (nIndex := 16#21A5, nSubIndex := 0); // Fixed 1 controller Ramp Time CoE register
    cRampMode_FIX1 : ST_CoEIndSub := (nIndex := 16#21A6, nSubIndex := 0); // Fixed 1 controller Ramp Mode CoE register
    cCtrlDir_FIX1 : ST_CoEIndSub := (nIndex := 16#21A7, nSubIndex := 0); // Fixed 1 controller Control Direction CoE register
    cPGain_FIX1 : ST_CoEIndSub := (nIndex := 16#21A8, nSubIndex := 0); // Fixed 1 controller P Gain CoE register
    cIGain_FIX1 : ST_CoEIndSub := (nIndex := 16#21A9, nSubIndex := 0); // Fixed 1 controller I Gain CoE register
    cRampTime_FIX2 : ST_CoEIndSub := (nIndex := 16#21AF, nSubIndex := 0); // Fixed 2 controller Ramp Time CoE register
    cRampMode_FIX2 : ST_CoEIndSub := (nIndex := 16#21B0, nSubIndex := 0); // Fixed 2 controller Ramp Mode CoE register
    cCtrlDir_FIX2 : ST_CoEIndSub := (nIndex := 16#21B1, nSubIndex := 0); // Fixed 2 controller Control Direction CoE register
    cPGain_FIX2 : ST_CoEIndSub := (nIndex := 16#21B2, nSubIndex := 0); // Fixed 2 controller P Gain CoE register
    cIGain_FIX2 : ST_CoEIndSub := (nIndex := 16#21B3, nSubIndex := 0); // Fixed 2 controller I Gain CoE register
    cRampTime_SP : ST_CoEIndSub := (nIndex := 16#21B9, nSubIndex := 0); // Soft Pump controller Ramp Time CoE register
    cRampMode_SP : ST_CoEIndSub := (nIndex := 16#21BA, nSubIndex := 0); // Soft Pump controller Ramp Time CoE register
    cPGain_SP : ST_CoEIndSub := (nIndex := 16#21BC, nSubIndex := 0); // Soft Pump controller Ramp Time CoE register
    cPosLimitOpen : ST_CoEIndSub := (nIndex := 16#56B3, nSubIndex := 0); // General open limit. It overides the PosLimitOpenCtrl if SET lower
    cPosLimitOpenCtrl : ST_CoEIndSub := (nIndex := 16#56B4, nSubIndex := 0); // Open limit active during pressure control only
END_VAR
VAR
    fCalcPosSP : REAL := 0;
    fCalcPresSP : REAL := 0;
    fPressRaw : REAL := 0;             // Ranges 0 to 1000000 (or 0.0 to 10V) (1E-12 to 1E-2)
    eValveModeSP : E_ControlModeSP;    // Control Mode setpoint internal variable
    fReqPos : REAL;                    // Requested position internal variable
    fReqPres : REAL;                   // Requested pressure internal variable

    bRemAcsToggle : BOOL;              // Remote access control bit
    //timer for zero function
    tZeroTogg : TON := (PT := T#1S);
    //timer for remote function
    tRemAcsTogg : TON := (PT := T#500MS);
    //used for logging
    ePreviousState : E_VCN_VAT590;

    (*CoE Interface*)
    (*Link this to your VAT590 reference variables under InfoData.*)
    //Connect i_stVat590PlcDriveRef.aNetId to the VAT590 Valve InfoData^AdsAddr^netId
    //Connect i_stVat590PlcDriveRef.nSlaveAddr to the VAT590 Valve InfoData^AdsAddr^port
    i_stVat590PlcDriveRef AT %I*: ST_PlcDriveRef;
    stVat590DriveRef : ST_DriveRef;

    fbCoeRead : FB_CoERead_ByDriveRef;   // CoE Read function block
    fbCoeWrite : FB_CoEWrite_ByDriveRef; // CoE Write function block

    stCoeParamsInternal : ST_VAT590_COE;   // Internal storage of CoE parameters
    nCaseReadCoe : UINT := 1;          // Iterator for going through all CoE parameters
    rtCoeReset : R_TRIG;               // Rising edge trigger for reset CoE Interface error
    ftCoeReadBusy : F_TRIG;            // Falling edge trigger for CoE read new data
    ftCoeWriteBusy : F_TRIG;           // Falling edge trigger for CoE write data
    bFirstRead : BOOL := TRUE;         // FALSE after succesfull first readout of all CoE parameters

    (*VAT590 Ethercat IO Interface*)
    // Ethercat Interface Inputs
    i_nRawPosition       AT %I* : DINT;               // Position readback from the valve
    i_nRawPressure       AT %I* : DINT;               // Pressure readback from the valve
    i_eControlMode       AT %I* : E_ControlMode;      // Valve control mode readback
    i_eFatalError        AT %I* : E_FatalErrors;      // Valve Fatal Errors readback
    i_stGenStatus        AT %I* : ST_GeneralStatus;   // Valve General Status readback
    i_stGenWarnings      AT %I* : ST_GeneralWarnings; // Valve General Warnings readback
    i_stExtnWarnings     AT %I* : ST_ExtendedWarnings;// Valve Extended Warnings readback
    // Ethercat Interface Outputs
    o_nRawPositionSP     AT %Q* : DINT;               // Position setpoint
    o_nRawPressureSP     AT %Q* : DINT;               // Pressure setpoint
    o_nRawPressure       AT %Q* : DINT;               // Raw pressure output, eliminate need for external connection of AI, ranges 0 to 1000000 (or 0.0 to 10V) (1E-12 Torr to 1E-2 Torr)
    o_eCtrlModeSP        AT %Q* : E_ControlModeSP;    // Valve control mode setpoint
    o_stGenCtrlSP        AT %Q* : ST_GeneralControlSP;// General Control setpoint
    (*Ethercat Interface Status Check*)
    (*Link this to your VAT590 WcState variable under WcState*)
    i_bValveEthCatStatus AT %I* : BOOL := TRUE;
END_VAR
VAR PERSISTENT
    fUpperLimit	: REAL;                // Max position in % that can be requested
    fPresMaxLim : REAL;                // Max pressure in Torr that can be requested
    fPresRbMaxLim : REAL;              // Max pressure in Torr read by chamber gauge, valve will close above the pressure.
END_VAR

(* Needle valve control FB
J. Govednik 2021-11-22

This FB should be used as a low level control block.

It provides:
Valve position ceiling
Interlock
CoE Interface R/W

It could be used for:
Valve position/flow linearization
*)

(*Set Coe Interface, AmsNetID, Slave address etc*)
SetCoeInterface();

(*Read from EPICS and Valve Ethercat interface*)
ReadFromInput();

(*Checking which Control mode is selected and if valve's communication is OK*)
IF stVcnVat590.bValveEthCatStatus THEN //If valve is not connected or something is wrong with EtherCAT communication PLC will set this bit to 1
    fReqPos := 0; //set req. position to 0
    eValveModeSP := E_ControlModeSP.CloseValve; //set control mode of the valve to CLOSE VALVE
    stVcnVat590.eValveControl := E_VCN_VAT590.CloseValve; //EPICS command hold in CloseValve state
    stVcnVat590.stValveStatus.eControlMode := E_ControlMode.FatalError; //override the readback from the valve because when valve is disconnected the value remains
    stVcnVat590.nRawPosition := 0; //override the readback from the valve because when valve is disconnected the value remains
    stVcnVat590.nRawPressure := 0; //override the readback from the valve because when valve is disconnected the value remains
ELSIF bExtIlkOK THEN
    CASE stVcnVat590.eValveControl OF
        E_VCN_VAT590.OpenValve:
            eValveModeSP := E_ControlModeSP.OpenValve;
        E_VCN_VAT590.CloseValve:
            eValveModeSP := E_ControlModeSP.CloseValve;
        E_VCN_VAT590.ManualControl:
            IF IG.xPRESS_OK AND IG.rPRESS <= fPresRbMaxLim THEN
                eValveModeSP := E_ControlModeSP.ManualControl;
            ELSE
                eValveModeSP := E_ControlModeSP.CloseValve; // Close valve if something is wrong with the gauge
                stVcnVat590.eValveControl := E_VCN_VAT590.CloseValve;
            END_IF
        E_VCN_VAT590.PressureControl:
            IF IG.xPRESS_OK AND IG.rPRESS <= fPresRbMaxLim THEN
                eValveModeSP := E_ControlModeSP.PressureControl;
            ELSE
                eValveModeSP := E_ControlModeSP.CloseValve; // Close valve if something is wrong with the gauge
                stVcnVat590.eValveControl := E_VCN_VAT590.CloseValve;
            END_IF
        E_VCN_VAT590.HoldValve:
            IF stVcnVat590.stValveStatus.eControlMode = E_ControlMode.ManualControl OR
                stVcnVat590.stValveStatus.eControlMode = E_ControlMode.PressureControl THEN
                eValveModeSP := E_ControlModeSP.HoldValve;
            END_IF
    END_CASE
ELSE
    fReqPos := 0;
    eValveModeSP := E_ControlModeSP.CloseValve;
    stVcnVat590.eValveControl := E_VCN_VAT590.CloseValve;
END_IF

(*Position SP calculation*)
fReqPos := LIMIT(0, fReqPos, fUpperLimit);
fCalcPosSP := fReqPos * (cOpenPosition-cClosePosition)/100 + cClosePosition;
fCalcPosSP := LIMIT(cClosePosition, fCalcPosSP, cOpenPosition); //The requested position SP should remain within this range

(*Pressure SP calculation*)
//Limit the input from EPICS between upper and lower limit defined for seleceted pressure sensor
fReqPres := LIMIT(cMinPress, fReqPres, fPresMaxLim);
//Calcuate pressure setpoint
fCalcPresSP := cPressRawSlope * LOG(fReqPres/cBasePress) + cPressRawBase;
fCalcPresSP := LIMIT(cPresSPLowLim, fCalcPresSP, cPresSPUpLim); //The requested pressure SP should remain within this range

(*Calculated Pressure SP, Pressure readback and PressureRaw output value are 0 if Pressure sensor is not working*)
//Calculate PressureRaw value linked to the Valve's External Digital pressure sensor 1 input
//Pressure information from IG input is linked to stVcnVat590.fPressure
IF IG.xPRESS_OK THEN
    stVcnVat590.fPressure := IG.rPRESS;
    fPressRaw := cPressRawSlope * LOG(IG.rPRESS/cBasePress) + cPressRawBase;
ELSE
    fCalcPresSP := 0;
    stVcnVat590.fPressure := 0;
    fPressRaw := 0;
END_IF

(*Zero function*)
IF stVcnVat590.stValveStatus.bZeroDisabled OR tZeroTogg.Q THEN
    stVcnVat590.bZero := FALSE;
END_IF
tZeroTogg.IN := stVcnVat590.bZero;
tZeroTogg();

(*Set Remote Access*)
IF stVcnVat590.stValveStatus.eRemoteStatus <> stVcnVat590.eRemoteControl THEN
    tRemAcsTogg.IN := TRUE;
    IF tRemAcsTogg.Q THEN
        bRemAcsToggle := NOT bRemAcsToggle;
        tRemAcsTogg.IN := FALSE;
    END_IF
END_IF
tRemAcsTogg();

(*Reset Coe Interface error*)
rtCoeReset(CLK := stVcnVat590.bResetCoeError);
IF rtCoeReset.Q THEN
    stVcnVat590.bResetCoeError := FALSE;
END_IF

(*Write CoE Parameters*)
WriteCoeParameters();

(*Read CoE Parameters*)
ReadCoeParameters();

(*Write to EPICS and Valve Ethercat interface*)
WriteToOutput();

(*Load or save the persistent variables*)
LoadPersistentData();

(*Logging*)
Logger();

ACTION LoadPersistentData:
(*On first PLC pass, load the persistent value into the structrue variable*)
IF (bRestorePersistentData) THEN
    bRestorePersistentData	:= FALSE;
    IF (fUpperLimit <> 0) THEN
        stVcnVat590.fPosSetLimit := fUpperLimit;
    END_IF;
    IF (fPresMaxLim <> 0) THEN
        stVcnVat590.fPresSetLimit := fPresMaxLim;
    END_IF;
    IF (fPresRbMaxLim <> 0) THEN
        stVcnVat590.fPresRdbkLimit := fPresRbMaxLim;
    END_IF;
END_IF
END_ACTION

ACTION Logger:
// ILK logger
IF NOT (stVcnVat590.bIlkOK ) AND NOT(ePreviousState = E_VCN_VAT590.CloseValve) THEN
         fbLogger(sMsg:='Lost interlock ok bit while valve was open.', eSevr:=TcEventSeverity.Critical);
END_IF


//Control STATE Logger
IF ePreviousState <> stVcnVat590.eValveControl THEN
      CASE stVcnVat590.eValveControl OF
        E_VCN_VAT590.ManualControl:
            fbLogger(sMsg:='Valve in manual control mode.', eSevr:=TcEventSeverity.Warning);
        E_VCN_VAT590.HoldValve:
            fbLogger(sMsg:='Valve in hold control mode.', eSevr:=TcEventSeverity.Warning);
        E_VCN_VAT590.OpenValve:
            fbLogger(sMsg:='Valve Open.', eSevr:=TcEventSeverity.Info);
        E_VCN_VAT590.PressureControl:
            fbLogger(sMsg:='Valve in pressure control mode.', eSevr:=TcEventSeverity.Info);
        E_VCN_VAT590.CloseValve:
            fbLogger(sMsg:='Valve closed.', eSevr:=TcEventSeverity.Info);
      END_CASE
      ePreviousState := stVcnVat590.eValveControl;
  END_IF


// Log valve open
tAction(CLK:= (stVcnVat590.eValveControl = E_VCN_VAT590.OpenValve) );
IF tAction.Q THEN fbLogger(sMsg:='Valve commanded to fully open', eSevr:=TcEventSeverity.Info); END_IF
END_ACTION

ACTION ReadCoeParameters:
CASE nCaseReadCoe OF
    0:
        stVcnVat590.bCoeError := TRUE;
        IF rtCoeReset.Q THEN
            nCaseReadCoe := 1;
            stVcnVat590.bCoeError := FALSE;
            bFirstRead := TRUE; // Set bFirstRead after Coe interface reset
        END_IF
    1:
        fbCoeRead.nIndex := cPressCtrl.nIndex;
        fbCoeRead.nSubIndex := cPressCtrl.nSubIndex;
        fbCoeRead.pDstBuf := ADR(stVcnVat590.stCoeParameters.ePIDCtrl);
        fbCoeRead.cbBufLen := SIZEOF(stVcnVat590.stCoeParameters.ePIDCtrl);
        fbCoeRead.bExecute := TRUE;
    2:
        fbCoeRead.nIndex := cSensorDelay_AD.nIndex;
        fbCoeRead.nSubIndex := cSensorDelay_AD.nSubIndex;
        fbCoeRead.pDstBuf := ADR(stVcnVat590.stCoeParameters.fSensorDelay_AD);
        fbCoeRead.cbBufLen := SIZEOF(stVcnVat590.stCoeParameters.fSensorDelay_AD);
        fbCoeRead.bExecute := TRUE;
    3:
        fbCoeRead.nIndex := cRampTime_AD.nIndex;
        fbCoeRead.nSubIndex := cRampTime_AD.nSubIndex;
        fbCoeRead.pDstBuf := ADR(stVcnVat590.stCoeParameters.fRampTime_AD);
        fbCoeRead.cbBufLen := SIZEOF(stVcnVat590.stCoeParameters.fRampTime_AD);
        fbCoeRead.bExecute := TRUE;
    4:
        fbCoeRead.nIndex := cRampMode_AD.nIndex;
        fbCoeRead.nSubIndex := cRampMode_AD.nSubIndex;
        fbCoeRead.pDstBuf := ADR(stVcnVat590.stCoeParameters.bRampMode_AD);
        fbCoeRead.cbBufLen := SIZEOF(stVcnVat590.stCoeParameters.bRampMode_AD);
        fbCoeRead.bExecute := TRUE;
    5:
        fbCoeRead.nIndex := cGainFactor_AD.nIndex;
        fbCoeRead.nSubIndex := cGainFactor_AD.nSubIndex;
        fbCoeRead.pDstBuf := ADR(stVcnVat590.stCoeParameters.fGainFactor_AD);
        fbCoeRead.cbBufLen := SIZEOF(stVcnVat590.stCoeParameters.fGainFactor_AD);
        fbCoeRead.bExecute := TRUE;
    6:
        fbCoeRead.nIndex := cRampTime_FIX1.nIndex;
        fbCoeRead.nSubIndex := cRampTime_FIX1.nSubIndex;
        fbCoeRead.pDstBuf := ADR(stVcnVat590.stCoeParameters.fRampTime_FIX1);
        fbCoeRead.cbBufLen := SIZEOF(stVcnVat590.stCoeParameters.fRampTime_FIX1);
        fbCoeRead.bExecute := TRUE;
    7:
        fbCoeRead.nIndex := cRampMode_FIX1.nIndex;
        fbCoeRead.nSubIndex := cRampMode_FIX1.nSubIndex;
        fbCoeRead.pDstBuf := ADR(stVcnVat590.stCoeParameters.bRampMode_FIX1);
        fbCoeRead.cbBufLen := SIZEOF(stVcnVat590.stCoeParameters.bRampMode_FIX1);
        fbCoeRead.bExecute := TRUE;
    8:
        fbCoeRead.nIndex := cCtrlDir_FIX1.nIndex;
        fbCoeRead.nSubIndex := cCtrlDir_FIX1.nSubIndex;
        fbCoeRead.pDstBuf := ADR(stVcnVat590.stCoeParameters.bCtrlDir_FIX1);
        fbCoeRead.cbBufLen := SIZEOF(stVcnVat590.stCoeParameters.bCtrlDir_FIX1);
        fbCoeRead.bExecute := TRUE;
    9:
        fbCoeRead.nIndex := cPGain_FIX1.nIndex;
        fbCoeRead.nSubIndex := cPGain_FIX1.nSubIndex;
        fbCoeRead.pDstBuf := ADR(stVcnVat590.stCoeParameters.fPGain_FIX1);
        fbCoeRead.cbBufLen := SIZEOF(stVcnVat590.stCoeParameters.fPGain_FIX1);
        fbCoeRead.bExecute := TRUE;
    10:
        fbCoeRead.nIndex := cIGain_FIX1.nIndex;
        fbCoeRead.nSubIndex := cIGain_FIX1.nSubIndex;
        fbCoeRead.pDstBuf := ADR(stVcnVat590.stCoeParameters.fIGain_FIX1);
        fbCoeRead.cbBufLen := SIZEOF(stVcnVat590.stCoeParameters.fIGain_FIX1);
        fbCoeRead.bExecute := TRUE;
    11:
        fbCoeRead.nIndex := cRampTime_FIX2.nIndex;
        fbCoeRead.nSubIndex := cRampTime_FIX2.nSubIndex;
        fbCoeRead.pDstBuf := ADR(stVcnVat590.stCoeParameters.fRampTime_FIX2);
        fbCoeRead.cbBufLen := SIZEOF(stVcnVat590.stCoeParameters.fRampTime_FIX2);
        fbCoeRead.bExecute := TRUE;
    12:
        fbCoeRead.nIndex := cRampMode_FIX2.nIndex;
        fbCoeRead.nSubIndex := cRampMode_FIX2.nSubIndex;
        fbCoeRead.pDstBuf := ADR(stVcnVat590.stCoeParameters.bRampMode_FIX2);
        fbCoeRead.cbBufLen := SIZEOF(stVcnVat590.stCoeParameters.bRampMode_FIX2);
        fbCoeRead.bExecute := TRUE;
    13:
        fbCoeRead.nIndex := cCtrlDir_FIX2.nIndex;
        fbCoeRead.nSubIndex := cCtrlDir_FIX2.nSubIndex;
        fbCoeRead.pDstBuf := ADR(stVcnVat590.stCoeParameters.bCtrlDir_FIX2);
        fbCoeRead.cbBufLen := SIZEOF(stVcnVat590.stCoeParameters.bCtrlDir_FIX2);
        fbCoeRead.bExecute := TRUE;
    14:
        fbCoeRead.nIndex := cPGain_FIX2.nIndex;
        fbCoeRead.nSubIndex := cPGain_FIX2.nSubIndex;
        fbCoeRead.pDstBuf := ADR(stVcnVat590.stCoeParameters.fPGain_FIX2);
        fbCoeRead.cbBufLen := SIZEOF(stVcnVat590.stCoeParameters.fPGain_FIX2);
        fbCoeRead.bExecute := TRUE;
    15:
        fbCoeRead.nIndex := cIGain_FIX2.nIndex;
        fbCoeRead.nSubIndex := cIGain_FIX2.nSubIndex;
        fbCoeRead.pDstBuf := ADR(stVcnVat590.stCoeParameters.fIGain_FIX2);
        fbCoeRead.cbBufLen := SIZEOF(stVcnVat590.stCoeParameters.fIGain_FIX2);
        fbCoeRead.bExecute := TRUE;
    16:
        fbCoeRead.nIndex := cRampTime_SP.nIndex;
        fbCoeRead.nSubIndex := cRampTime_SP.nSubIndex;
        fbCoeRead.pDstBuf := ADR(stVcnVat590.stCoeParameters.fRampTime_SP);
        fbCoeRead.cbBufLen := SIZEOF(stVcnVat590.stCoeParameters.fRampTime_SP);
        fbCoeRead.bExecute := TRUE;
    17:
        fbCoeRead.nIndex := cRampMode_SP.nIndex;
        fbCoeRead.nSubIndex := cRampMode_SP.nSubIndex;
        fbCoeRead.pDstBuf := ADR(stVcnVat590.stCoeParameters.bRampMode_SP);
        fbCoeRead.cbBufLen := SIZEOF(stVcnVat590.stCoeParameters.bRampMode_SP);
        fbCoeRead.bExecute := TRUE;
    18:
        fbCoeRead.nIndex := cPGain_SP.nIndex;
        fbCoeRead.nSubIndex := cPGain_SP.nSubIndex;
        fbCoeRead.pDstBuf := ADR(stVcnVat590.stCoeParameters.fPGain_SP);
        fbCoeRead.cbBufLen := SIZEOF(stVcnVat590.stCoeParameters.fPGain_SP);
        fbCoeRead.bExecute := TRUE;
    19:
        fbCoeRead.nIndex := cPosLimitOpen.nIndex;
        fbCoeRead.nSubIndex := cPosLimitOpen.nSubIndex;
        fbCoeRead.pDstBuf := ADR(stVcnVat590.stCoeParameters.fPositionLimitOpen);
        fbCoeRead.cbBufLen := SIZEOF(stVcnVat590.stCoeParameters.fPositionLimitOpen);
        fbCoeRead.bExecute := TRUE;
    20:
        fbCoeRead.nIndex := cPosLimitOpenCtrl.nIndex;
        fbCoeRead.nSubIndex := cPosLimitOpenCtrl.nSubIndex;
        fbCoeRead.pDstBuf := ADR(stVcnVat590.stCoeParameters.fPositionLimitOpenControl);
        fbCoeRead.cbBufLen := SIZEOF(stVcnVat590.stCoeParameters.fPositionLimitOpenControl);
        fbCoeRead.bExecute := TRUE;
END_CASE

ftCoeReadBusy(CLK:=fbCoeRead.bBusy);
IF ftCoeReadBusy.Q THEN
    fbCoeRead.bExecute := FALSE;
    IF NOT fbCoeRead.bError THEN
        nCaseReadCoe := nCaseReadCoe + 1;
        IF nCaseReadCoe > 20 THEN
            nCaseReadCoe := 1;
            bFirstRead := FALSE; // Reset bFirstRead after successfull readout of all parameters
        END_IF
    ELSE
        nCaseReadCoe := 0; // Go to Error state
    END_IF
END_IF

fbCoeRead();
stCoeParamsInternal := stVcnVat590.stCoeParameters; //Save current values to internal structure
END_ACTION

ACTION ReadFromInput:
(*Read from EPICS*)
fUpperLimit := LIMIT(0, stVcnVat590.fPosSetLimit, 100);
fPresMaxLim := LIMIT(cMinPress, stVcnVat590.fPresSetLimit, cMaxPress);
fPresRbMaxLim := LIMIT(cMinPress, stVcnVat590.fPresRdbkLimit, cMaxPress);
fReqPos := LIMIT(0, stVcnVat590.fReqPosition, 100);
fReqPres := LIMIT(cMinPress, stVcnVat590.fReqPressure, cMaxPress);

(*Read from VAT valve*)
stVcnVat590.stValveStatus.eControlMode := i_eControlMode;
stVcnVat590.stValveStatus.eFatalErrors := i_eFatalError;
stVcnVat590.nRawPosition := i_nRawPosition;
stVcnVat590.nRawPressure := i_nRawPressure;
//Mapping General statuses
stVcnVat590.stValveStatus.bFieldBusDatavalid := i_stGenStatus.Bit0FieldBusDatavalid;
stVcnVat590.stValveStatus.bZeroExecuted := i_stGenStatus.Bit1ZeroExecuted;
stVcnVat590.stValveStatus.bPingPongRxBit := i_stGenStatus.Bit2PingPongRxBit;
stVcnVat590.stValveStatus.bPressureSimulation := i_stGenStatus.Bit3PressureSimulation;
stVcnVat590.stValveStatus.bPressureSPReached := i_stGenStatus.Bit4PressureSPReached;
stVcnVat590.stValveStatus.bWarningsActive := i_stGenStatus.Bit9WarningsActive;
//Read Remote status
stVcnVat590.stValveStatus.eRemoteStatus.0 := i_stGenStatus.Bit7AccessModeBit0;
stVcnVat590.stValveStatus.eRemoteStatus.1 := i_stGenStatus.Bit8AccessModeBit1;
//Mapping General warnings
stVcnVat590.stValveStatus.bServiceRequest := i_stGenWarnings.Bit0ServiceRequest;
stVcnVat590.stValveStatus.bPowerFailureBattery := i_stGenWarnings.Bit3PowerFailureBattery;
stVcnVat590.stValveStatus.bSensMeasUnitFault := i_stGenWarnings.Bit10SensMeasUnitFault;
//Mapping Extended warnings
stVcnVat590.stValveStatus.bRemoteControlNotPossible := i_stExtnWarnings.Bit0RemoteControlNotPossible;
stVcnVat590.stValveStatus.bControlModeSPNotAllowed := i_stExtnWarnings.Bit1ControlModeSPNotAllowed;
stVcnVat590.stValveStatus.bZeroDisabled := i_stExtnWarnings.Bit2ZeroDisabled;
stVcnVat590.stValveStatus.bPFODeactivated := i_stExtnWarnings.Bit3PFODeactivated;
stVcnVat590.stValveStatus.bPressureSPOutOfRange := i_stExtnWarnings.Bit5PressureSPOutOfRange;
stVcnVat590.stValveStatus.bPositionSPOutOfRange := i_stExtnWarnings.Bit6PositionSPOutOfRange;
stVcnVat590.stValveStatus.bCtrlSPOutOfRange := i_stExtnWarnings.Bit10CtrlSPOutOfRange;
stVcnVat590.stValveStatus.bGeneralCtrlSPOutOfRange := i_stExtnWarnings.Bit11GeneralCtrlSPOutOfRange;
stVcnVat590.stValveStatus.bProcDataSettingsNotvalid := i_stExtnWarnings.Bit12ProcDataSettingsNotvalid;
//Mapping WcState - Valve Ethercat Status
stVcnVat590.bValveEthCatStatus := i_bValveEthCatStatus;
END_ACTION

ACTION SetCoeInterface:
stVat590DriveRef.sNetId := F_CreateAmsNetId(i_stVat590PlcDriveRef.aNetId);
stVat590DriveRef.nSlaveAddr := i_stVat590PlcDriveRef.nSlaveAddr;
stVat590DriveRef.nDriveNo := i_stVat590PlcDriveRef.nDriveNo;
stVat590DriveRef.nDriveType := i_stVat590PlcDriveRef.nDriveType;
fbCoeRead.stDriveRef := stVat590DriveRef;
fbCoeWrite.stDriveRef := stVat590DriveRef;
END_ACTION

METHOD SetThrottle : BOOL
VAR_INPUT
    rUpperLimit	:	REAL;
END_VAR
stVcnVat590.fPosSetLimit := LIMIT(0, rUpperLimit, 100);
END_METHOD

METHOD ValveControl : BOOL
VAR_INPUT
    state : E_VCN_VAT590; // Set Control modes
END_VAR
stVcnVat590.eValveControl := state;
END_METHOD

ACTION WriteCoeParameters:
// User will change one parameter at a time so solution with ELSIF should work OK
IF stVcnVat590.bCoeError THEN
    IF rtCoeReset.Q THEN
        stVcnVat590.bCoeError := FALSE;
    END_IF;
ELSIF bFirstRead THEN
    ;//Wait until first readout of all CoE parameters is completed
ELSIF stVcnVat590.stCoeParameters.ePIDCtrl <> stCoeParamsInternal.ePIDCtrl THEN
    fbCoeWrite.nIndex := cPressCtrl.nIndex;
    fbCoeWrite.nSubIndex := cPressCtrl.nSubIndex;
    fbCoeWrite.pSrcBuf := ADR(stVcnVat590.stCoeParameters.ePIDCtrl);
    fbCoeWrite.cbBufLen := SIZEOF(stVcnVat590.stCoeParameters.ePIDCtrl);
    fbCoeWrite.bExecute := TRUE;
ELSIF stVcnVat590.stCoeParameters.fSensorDelay_AD <> stCoeParamsInternal.fSensorDelay_AD THEN
    fbCoeWrite.nIndex := cSensorDelay_AD.nIndex;
    fbCoeWrite.nSubIndex := cSensorDelay_AD.nSubIndex;
    fbCoeWrite.pSrcBuf := ADR(stVcnVat590.stCoeParameters.fSensorDelay_AD);
    fbCoeWrite.cbBufLen := SIZEOF(stVcnVat590.stCoeParameters.fSensorDelay_AD);
    fbCoeWrite.bExecute := TRUE;
ELSIF stVcnVat590.stCoeParameters.fRampTime_AD <> stCoeParamsInternal.fRampTime_AD THEN
    fbCoeWrite.nIndex := cRampTime_AD.nIndex;
    fbCoeWrite.nSubIndex := cRampTime_AD.nSubIndex;
    fbCoeWrite.pSrcBuf := ADR(stVcnVat590.stCoeParameters.fRampTime_AD);
    fbCoeWrite.cbBufLen := SIZEOF(stVcnVat590.stCoeParameters.fRampTime_AD);
    fbCoeWrite.bExecute := TRUE;
ELSIF stVcnVat590.stCoeParameters.bRampMode_AD <> stCoeParamsInternal.bRampMode_AD THEN
    fbCoeWrite.nIndex := cRampMode_AD.nIndex;
    fbCoeWrite.nSubIndex := cRampMode_AD.nSubIndex;
    fbCoeWrite.pSrcBuf := ADR(stVcnVat590.stCoeParameters.bRampMode_AD);
    fbCoeWrite.cbBufLen := SIZEOF(stVcnVat590.stCoeParameters.bRampMode_AD);
    fbCoeWrite.bExecute := TRUE;
ELSIF stVcnVat590.stCoeParameters.fGainFactor_AD <> stCoeParamsInternal.fGainFactor_AD THEN
    fbCoeWrite.nIndex := cGainFactor_AD.nIndex;
    fbCoeWrite.nSubIndex := cGainFactor_AD.nSubIndex;
    fbCoeWrite.pSrcBuf := ADR(stVcnVat590.stCoeParameters.fGainFactor_AD);
    fbCoeWrite.cbBufLen := SIZEOF(stVcnVat590.stCoeParameters.fGainFactor_AD);
    fbCoeWrite.bExecute := TRUE;
ELSIF stVcnVat590.stCoeParameters.fRampTime_FIX1 <> stCoeParamsInternal.fRampTime_FIX1 THEN
    fbCoeWrite.nIndex := cRampTime_FIX1.nIndex;
    fbCoeWrite.nSubIndex := cRampTime_FIX1.nSubIndex;
    fbCoeWrite.pSrcBuf := ADR(stVcnVat590.stCoeParameters.fRampTime_FIX1);
    fbCoeWrite.cbBufLen := SIZEOF(stVcnVat590.stCoeParameters.fRampTime_FIX1);
    fbCoeWrite.bExecute := TRUE;
ELSIF stVcnVat590.stCoeParameters.bRampMode_FIX1 <> stCoeParamsInternal.bRampMode_FIX1 THEN
    fbCoeWrite.nIndex := cRampMode_FIX1.nIndex;
    fbCoeWrite.nSubIndex := cRampMode_FIX1.nSubIndex;
    fbCoeWrite.pSrcBuf := ADR(stVcnVat590.stCoeParameters.bRampMode_FIX1);
    fbCoeWrite.cbBufLen := SIZEOF(stVcnVat590.stCoeParameters.bRampMode_FIX1);
    fbCoeWrite.bExecute := TRUE;
ELSIF stVcnVat590.stCoeParameters.bCtrlDir_FIX1 <> stCoeParamsInternal.bCtrlDir_FIX1 THEN
    fbCoeWrite.nIndex := cCtrlDir_FIX1.nIndex;
    fbCoeWrite.nSubIndex := cCtrlDir_FIX1.nSubIndex;
    fbCoeWrite.pSrcBuf := ADR(stVcnVat590.stCoeParameters.bCtrlDir_FIX1);
    fbCoeWrite.cbBufLen := SIZEOF(stVcnVat590.stCoeParameters.bCtrlDir_FIX1);
    fbCoeWrite.bExecute := TRUE;
ELSIF stVcnVat590.stCoeParameters.fPGain_FIX1 <> stCoeParamsInternal.fPGain_FIX1 THEN
    fbCoeWrite.nIndex := cPGain_FIX1.nIndex;
    fbCoeWrite.nSubIndex := cPGain_FIX1.nSubIndex;
    fbCoeWrite.pSrcBuf := ADR(stVcnVat590.stCoeParameters.fPGain_FIX1);
    fbCoeWrite.cbBufLen := SIZEOF(stVcnVat590.stCoeParameters.fPGain_FIX1);
    fbCoeWrite.bExecute := TRUE;
ELSIF stVcnVat590.stCoeParameters.fIGain_FIX1 <> stCoeParamsInternal.fIGain_FIX1 THEN
    fbCoeWrite.nIndex := cIGain_FIX1.nIndex;
    fbCoeWrite.nSubIndex := cIGain_FIX1.nSubIndex;
    fbCoeWrite.pSrcBuf := ADR(stVcnVat590.stCoeParameters.fIGain_FIX1);
    fbCoeWrite.cbBufLen := SIZEOF(stVcnVat590.stCoeParameters.fIGain_FIX1);
    fbCoeWrite.bExecute := TRUE;
ELSIF stVcnVat590.stCoeParameters.fRampTime_FIX2 <> stCoeParamsInternal.fRampTime_FIX2 THEN
    fbCoeWrite.nIndex := cRampTime_FIX2.nIndex;
    fbCoeWrite.nSubIndex := cRampTime_FIX2.nSubIndex;
    fbCoeWrite.pSrcBuf := ADR(stVcnVat590.stCoeParameters.fRampTime_FIX2);
    fbCoeWrite.cbBufLen := SIZEOF(stVcnVat590.stCoeParameters.fRampTime_FIX2);
    fbCoeWrite.bExecute := TRUE;
ELSIF stVcnVat590.stCoeParameters.bRampMode_FIX2 <> stCoeParamsInternal.bRampMode_FIX2 THEN
    fbCoeWrite.nIndex := cRampMode_FIX2.nIndex;
    fbCoeWrite.nSubIndex := cRampMode_FIX2.nSubIndex;
    fbCoeWrite.pSrcBuf := ADR(stVcnVat590.stCoeParameters.bRampMode_FIX2);
    fbCoeWrite.cbBufLen := SIZEOF(stVcnVat590.stCoeParameters.bRampMode_FIX2);
    fbCoeWrite.bExecute := TRUE;
ELSIF stVcnVat590.stCoeParameters.bCtrlDir_FIX2 <> stCoeParamsInternal.bCtrlDir_FIX2 THEN
    fbCoeWrite.nIndex := cCtrlDir_FIX2.nIndex;
    fbCoeWrite.nSubIndex := cCtrlDir_FIX2.nSubIndex;
    fbCoeWrite.pSrcBuf := ADR(stVcnVat590.stCoeParameters.bCtrlDir_FIX2);
    fbCoeWrite.cbBufLen := SIZEOF(stVcnVat590.stCoeParameters.bCtrlDir_FIX2);
    fbCoeWrite.bExecute := TRUE;
ELSIF stVcnVat590.stCoeParameters.fPGain_FIX2 <> stCoeParamsInternal.fPGain_FIX2 THEN
    fbCoeWrite.nIndex := cPGain_FIX2.nIndex;
    fbCoeWrite.nSubIndex := cPGain_FIX2.nSubIndex;
    fbCoeWrite.pSrcBuf := ADR(stVcnVat590.stCoeParameters.fPGain_FIX2);
    fbCoeWrite.cbBufLen := SIZEOF(stVcnVat590.stCoeParameters.fPGain_FIX2);
    fbCoeWrite.bExecute := TRUE;
ELSIF stVcnVat590.stCoeParameters.fIGain_FIX2 <> stCoeParamsInternal.fIGain_FIX2 THEN
    fbCoeWrite.nIndex := cIGain_FIX2.nIndex;
    fbCoeWrite.nSubIndex := cIGain_FIX2.nSubIndex;
    fbCoeWrite.pSrcBuf := ADR(stVcnVat590.stCoeParameters.fIGain_FIX2);
    fbCoeWrite.cbBufLen := SIZEOF(stVcnVat590.stCoeParameters.fIGain_FIX2);
    fbCoeWrite.bExecute := TRUE;
ELSIF stVcnVat590.stCoeParameters.fRampTime_SP <> stCoeParamsInternal.fRampTime_SP THEN
    fbCoeWrite.nIndex := cRampTime_SP.nIndex;
    fbCoeWrite.nSubIndex := cRampTime_SP.nSubIndex;
    fbCoeWrite.pSrcBuf := ADR(stVcnVat590.stCoeParameters.fRampTime_SP);
    fbCoeWrite.cbBufLen := SIZEOF(stVcnVat590.stCoeParameters.fRampTime_SP);
    fbCoeWrite.bExecute := TRUE;
ELSIF stVcnVat590.stCoeParameters.bRampMode_SP <> stCoeParamsInternal.bRampMode_SP THEN
    fbCoeWrite.nIndex := cRampMode_SP.nIndex;
    fbCoeWrite.nSubIndex := cRampMode_SP.nSubIndex;
    fbCoeWrite.pSrcBuf := ADR(stVcnVat590.stCoeParameters.bRampMode_SP);
    fbCoeWrite.cbBufLen := SIZEOF(stVcnVat590.stCoeParameters.bRampMode_SP);
    fbCoeWrite.bExecute := TRUE;
ELSIF stVcnVat590.stCoeParameters.fPGain_SP <> stCoeParamsInternal.fPGain_SP THEN
    fbCoeWrite.nIndex := cPGain_SP.nIndex;
    fbCoeWrite.nSubIndex := cPGain_SP.nSubIndex;
    fbCoeWrite.pSrcBuf := ADR(stVcnVat590.stCoeParameters.fPGain_SP);
    fbCoeWrite.cbBufLen := SIZEOF(stVcnVat590.stCoeParameters.fPGain_SP);
    fbCoeWrite.bExecute := TRUE;
ELSIF stVcnVat590.stCoeParameters.fPositionLimitOpen <> stCoeParamsInternal.fPositionLimitOpen THEN
    fbCoeWrite.nIndex := cPosLimitOpen.nIndex;
    fbCoeWrite.nSubIndex := cPosLimitOpen.nSubIndex;
    fbCoeWrite.pSrcBuf := ADR(stVcnVat590.stCoeParameters.fPositionLimitOpen);
    fbCoeWrite.cbBufLen := SIZEOF(stVcnVat590.stCoeParameters.fPositionLimitOpen);
    fbCoeWrite.bExecute := TRUE;
ELSIF stVcnVat590.stCoeParameters.fPositionLimitOpenControl <> stCoeParamsInternal.fPositionLimitOpenControl THEN
    fbCoeWrite.nIndex := cPosLimitOpenCtrl.nIndex;
    fbCoeWrite.nSubIndex := cPosLimitOpenCtrl.nSubIndex;
    fbCoeWrite.pSrcBuf := ADR(stVcnVat590.stCoeParameters.fPositionLimitOpenControl);
    fbCoeWrite.cbBufLen := SIZEOF(stVcnVat590.stCoeParameters.fPositionLimitOpenControl);
    fbCoeWrite.bExecute := TRUE;
END_IF

ftCoeWriteBusy(CLK:=fbCoeWrite.bBusy);
IF ftCoeWriteBusy.Q THEN
    fbCoeWrite.bExecute := FALSE;
    IF fbCoeWrite.bError THEN
        stVcnVat590.bCoeError := TRUE;
    END_IF
END_IF

fbCoeWrite();
END_ACTION

ACTION WriteToOutput:
(*Write to EPICS*)
stVcnVat590.bIlkOK := bExtIlkOK;
stVcnVat590.nPositionSP := REAL_TO_DINT(fCalcPosSP);
stVcnVat590.nPressureSP := REAL_TO_DINT(fCalcPresSP);
stVcnVat590.fReqPosition := fReqPos;
stVcnVat590.fReqPressure := fReqPres;
stVcnVat590.fPresSetLimit := fPresMaxLim;
stVcnVat590.fPosSetLimit := fUpperLimit;

(*Write to VAT valve*)
o_eCtrlModeSP := eValveModeSP;
o_nRawPositionSP := REAL_TO_DINT(fCalcPosSP);
o_nRawPressureSP := REAL_TO_DINT(fCalcPresSP);
o_nRawPressure := REAL_TO_DINT(fPressRaw);
o_stGenCtrlSP.Bit0ExecuteZero := stVcnVat590.bZero;
o_stGenCtrlSP.Bit4AccessMode := bRemAcsToggle;
END_ACTION

END_FUNCTION_BLOCK

// ---- POUs/Functions/Valves/FB_VFS.TcPOU
(* This function block implements basic functionality for Fast Shutter/Valves*)
(* Create a separate virtual PLC for the fast shutter logic, and tie/map this task to the FAST I/O portion of the ethercat bus,
 so we can scan these I/Os faster than the rest of the vacuum I/Os.
The Fast shutter was tested with PLC task Cycle Base Time 50us with cycle time 0.050ms.
*)
FUNCTION_BLOCK FB_VFS EXTENDS FB_Valve
VAR_INPUT
    i_xPMPS_OK:	BOOL	; (*External MPS interlock, Set to TRUE when no PMPS interlock is required*)
    i_xExt_OK: BOOL; (*Other External Interlock, Set to True when no external interlock is required*)
    i_sDevName : T_MaxString :=  'VGC'; // Device name for diagnostic
    i_xVeto_Enable:BOOL:= FALSE; (*Set to TRUE if there is a Veto Valve to this VFS*)
END_VAR
VAR_IN_OUT
    io_fbFFHWO    :    FB_HardwareFFOutput;
END_VAR
VAR
    xOPN_OK :BOOL;
    xERR_ExtFault :BOOL;
    xVeto: BOOL;
    // PMPS
    fbFF    :    FB_FastFault :=(
        i_DevName := 'VFS',
        i_Desc := 'Fault occurs when fast valve is not in open state',
        i_TypeCode := 16#1010);

    rDiffPressAllowed	:	REAL := 22.5; // Torr, Default value comes from Vat Valve Manual
    rDiffPress : REAL;
    set : BOOL;
    reset: BOOL;

    xFirstPass	:	BOOL := TRUE;
    //fbFSInit		:	R_TRIG;
    rtOPN_SW :	R_TRIG;

    tonDelOK : TON;
    rtOK	:	R_TRIG;
    tonOvrd	:	TON;

    tDelOK	:	TIME := T#60S;
    tOvrd	:	TIME := T#10s;
    rTrigOverrideOpen : R_TRIG;

    xClose: BOOL;
    xOpen: BOOL;
    CloseTimer: TON;
    TimDur: TIME := T#20MS;
    OpenTimer: TON;
    OpenTimDur: TIME := T#2S;

    (* Timeouts*)
    tCLSTimeOutDuration: TIME:= T#0.5S;
    tOPNTimeOutDuration: TIME:= T#10S;
    tOPNtimeout: TON;
    tCLStimeout:TON;


    (*IO*)
    i_xOpnLS	AT%I*: BOOL;
    i_xClsLS	AT%I*: BOOL;
    q_xClose_A	AT%Q*: BOOL;
    q_xClose_B	AT%Q*: BOOL;
    q_xClose_C	AT%Q*: BOOL;
    q_xOPN_DO	AT%Q*: BOOL;
    i_xTrigger	AT%I*: BOOL;

    (*VETO Devices*)
    i_xVetoValveOpenDO AT%I*: BOOL;
    i_xVetoValveClosed AT%I*: BOOL;

    // Interface
    i_xPress_OK AT%I*:BOOL; (*To be linked to the Fast sensor structure signal IG.xPRESS_OK, to make sure that the device is connected*)
    i_xOPN_SW AT%I*:BOOL;
    i_xCLS_SW AT%I*:BOOL; (*external open signal e.g epics*)
    i_xVAC_FAULT_Reset	AT%I*: BOOL;(*Valve Vacuum OK, is set to False when there is Vacuum Fault*)
    i_xOverrideMode AT%I*: BOOL; (*To be linked to global override bit. This Overrides Vacuum logic only, EPS, MPS and PMPS are still enforces*)
    i_xOverrideOpen AT%I*: BOOL;
    q_xTrigger	AT%Q*: BOOL; (*Interface*)
    q_xVFS_Open AT%Q*: BOOL; (*Interface*)
    q_xVFS_Closed AT%Q*: BOOL; (*Interface*)
    q_xVAC_FAULT_OK AT%Q*: BOOL; (*Valve Vacuum OK, is set to False when there is Vacuum Fault*)
    q_xMPS_OK	 AT%Q*:	BOOL; (*MPS Fault OK, is set when the Valve is Open and there is no trigger*)
    q_eVFS_State AT%Q*: E_VGC; (*Interface*)

END_VAR



(* Fast Shutter/Valve Function Block*)
(* M.Ghaly Feb 2019*)

